(* IEC 61131-3 sources: TBEN-L5-PLC-11/src/st, 44 files *)

(* ---- E_IolAccess.st ---- *)
{attribute 'qualified_only'}
// Quyền truy cập tham số theo IODD (accessRights)
TYPE E_IolAccess :
(
    RO := 0,
    WO := 1,
    RW := 2
) INT;
END_TYPE

(* ---- E_IolCallState.st ---- *)
{attribute 'qualified_only'}
// Trạng thái state machine IOL_CALL của FB_IolMaster
TYPE E_IolCallState :
(
    IDLE      := 0,   // rảnh, chờ request trong FIFO
    WRITE_REQ := 1,   // WRREC khung IOL_CALL vào record CAP 0xB400
    RETRY_WR  := 2,   // master báo bận -> chờ rồi ghi lại
    READ_WAIT := 3,   // REQ đã hạ, chờ trước khi RDREC phản hồi
    READ_REQ  := 4,   // RDREC đọc phản hồi + kiểm khung
    DONE      := 5,   // trả kết quả cho client (1 chu kỳ)
    ERROR     := 6,   // trả lỗi cho client (1 chu kỳ)
    TIMEOUT   := 7,   // quá hạn: hạ REQ, chờ transport hết BUSY
    STUCK     := 8    // transport kẹt BUSY > 1 s, chỉ thoát bằng xReset
) INT;
END_TYPE

(* ---- E_IolCallStep.st ---- *)
{attribute 'qualified_only'}
// Bước handshake của client FB_IolCall
TYPE E_IolCallStep :
(
    IDLE := 0,
    WAIT := 1,    // đã vào hàng đợi master, chờ kết quả
    DONE := 2,
    ERR  := 3
) INT;
END_TYPE

(* ---- E_IolDataType.st ---- *)
{attribute 'qualified_only'}
// Kiểu dữ liệu tham số theo IODD (giá trị trên dây là big-endian)
TYPE E_IolDataType :
(
    U8    := 0,
    U16   := 1,
    U32   := 2,
    I8    := 3,
    I16   := 4,
    I32   := 5,
    STR   := 6,
    OCTET := 7    // record nhiều trường, lớp con tự tách (vd Limit index 64)
) INT;
END_TYPE

(* ---- E_IolDevJob.st ---- *)
{attribute 'qualified_only'}
// Loại việc ISDU đang chạy trong FB_IolDevBase
TYPE E_IolDevJob :
(
    NONE     := 0,
    IDENT    := 1,  // đọc index 16..24
    PARAM_RD := 2,  // đọc 1 tham số trong bảng
    PARAM_WR := 3,  // ghi 1 tham số trong bảng
    CUSTOM   := 4   // ISDU tự do của lớp con (system command, event list...)
) INT;
END_TYPE

(* ---- E_IolDevSeq.st ---- *)
{attribute 'qualified_only'}
// Bước trình tự gọi ISDU trong FB_IolDevBase
TYPE E_IolDevSeq :
(
    IDLE    := 0,   // chọn việc tiếp theo
    RUN     := 1,   // FB_IolCall đang chạy
    RELEASE := 2    // hạ Execute, chờ FB_IolCall về IDLE
) INT;
END_TYPE

(* ---- E_IolErrSource.st ---- *)
{attribute 'qualified_only'}
// Nguồn lỗi của 1 lần gọi IO-Link, để HMI biết lỗi nằm ở tầng nào
TYPE E_IolErrSource :
(
    NONE         := 0,
    PNIO         := 1,    // RDREC/WRREC trả STATUS lỗi (hoặc transport chưa cấu hình)
    IOL_MASTER   := 2,    // AL1100 báo IOL_M_ErrorCode
    IOL_DEVICE   := 3,    // cảm biến báo lỗi ISDU 0x80xx
    TIMEOUT      := 4,
    PARAM        := 5,    // tham số yêu cầu sai, không gửi đi
    LOCK         := 6,    // hết chỗ hàng đợi / không đăng ký được / bị reset
    FRAME        := 7,    // khung phản hồi sai
    NO_DEVICE    := 8,    // PQI.DA = 0: port không có thiết bị
    WRITE_LOCKED := 9,    // ghi bị khoá (chưa bật xMaintEnable)
    RANGE        := 10    // giá trị đặt ngoài dải IODD, chặn trước khi gửi
) INT;
END_TYPE

(* ---- E_IolEvtType.st ---- *)
{attribute 'qualified_only'}
// Loại event IO-Link (= bit 5..4 của EventQualifier)
TYPE E_IolEvtType :
(
    NOTIFICATION := 1,
    WARNING      := 2,
    ERROR        := 3
) INT;
END_TYPE

(* ---- E_IolService.st ---- *)
{attribute 'qualified_only'}
// Giá trị byte Control của khung IOL_CALL (request)
TYPE E_IolService :
(
    WRITE := 2,   // ISDU write
    READ  := 3    // ISDU read
) USINT;
END_TYPE

(* ---- E_O5D150_Param.st ---- *)
{attribute 'qualified_only'}
// Vị trí tham số trong bảng GVL_O5D150_Def.aParamDef (không phải IO-Link index)
TYPE E_O5D150_Param :
(
    SP1       := 0,   // index 60 sub 1
    CFG_LOGIC := 1,   // index 61 sub 1
    LIMITS    := 2,   // index 64 (min, max) - không đặt tên LIMIT vì trùng hàm chuẩn
    ALIGN     := 3,   // index 69
    LASER     := 4,   // index 80
    DISPLAY   := 5,   // index 96
    KEYLOCK   := 6,   // index 100
    DFO       := 7,   // index 74
    DS        := 8,   // index 76
    DR        := 9    // index 78
) INT;
END_TYPE

(* ---- ST_HMI_O5D150.st ---- *)
// Giao tiếp HMI <-> FB_Dev_O5D150 (lệnh: HMI đặt TRUE, PRG_IOLink tự xoá)
TYPE ST_HMI_O5D150 :
STRUCT
    // --- Lệnh ---
    xCmdReadAll      : BOOL;
    xCmdReadIdent    : BOOL;
    xCmdWriteSP1     : BOOL;          // ghi uiSetSP1 (cần xMaintEnable)
    xCmdWriteLogic   : BOOL;
    xCmdWriteLaser   : BOOL;
    xCmdWriteDisplay : BOOL;
    xCmdTestEvt1On   : BOOL;          // System Command 240 (cần xMaintEnable)
    xCmdTestEvt1Off  : BOOL;          // 241
    xCmdTestEvt2On   : BOOL;          // 242
    xCmdTestEvt2Off  : BOOL;          // 243
    xCmdReadEvents   : BOOL;          // đọc index 37 ngay (thử lại cả khi đã báo không hỗ trợ)
    xCmdResetErr     : BOOL;
    xAlignMode       : BOOL;          // giữ TRUE: đọc Align (69) chu kỳ chậm

    // --- Giá trị đặt ---
    uiSetSP1         : UINT := 100;   // cm, 5..200
    usiSetLogic      : USINT;         // 0 NO, 1 NC
    usiSetLaser      : USINT := 1;    // 0 Off, 1 On
    usiSetDisplay    : USINT := 1;    // 0 Off, 1 On, 2 Rotated

    // --- Process data ---
    uiDistance_cm    : UINT;
    rDistance_m      : REAL;
    xOut1            : BOOL;
    xPdValid         : BOOL;
    xOutOfRange      : BOOL;
    xPQ              : BOOL;
    xDA              : BOOL;
    xDE              : BOOL;

    // --- Tham số đọc về ---
    uiSP1            : UINT;
    usiLogic         : USINT;
    uiLimitMin_cm    : UINT;
    uiLimitMax_cm    : UINT;
    usiAlign         : USINT;         // %
    usiLaser         : USINT;
    usiDisplay       : USINT;
    xParamValid      : BOOL;          // SP1 đọc được lần gần nhất

    // --- Nhận dạng ---
    sVendor          : STRING(64);
    sProduct         : STRING(64);
    sSerial          : STRING(64);
    sFwRev           : STRING(64);

    // --- Event ---
    axEvtActive      : ARRAY[0..GVL_O5D150_Def.iEVT_COUNT - 1] OF BOOL;   // theo GVL_O5D150_Def.aEvtDef
    uiEvtCount       : UINT;
    wUnknownEvt      : WORD;
    xEvtListNotSupported : BOOL;

    // --- Trạng thái / lỗi ---
    xBusy            : BOOL;
    xError           : BOOL;          // lỗi gần nhất (giữ tới xCmdResetErr)
    uiDevErr         : UINT;
    wsErrText        : WSTRING(80);
    xWriteLocked     : BOOL;          // = NOT xMaintEnable
END_STRUCT
END_TYPE

(* ---- ST_IolEventDef.st ---- *)
// Định nghĩa 1 event của device (từ IODD)
TYPE ST_IolEventDef :
STRUCT
    wCode  : WORD;
    sName  : STRING(12);        // tên ngắn trên màn hình cảm biến
    wsText : WSTRING(48);       // mô tả cho HMI
    eType  : E_IolEvtType;
END_STRUCT
END_TYPE

(* ---- ST_IolIdent.st ---- *)
// Thông tin nhận dạng chuẩn IO-Link (index 16..24)
TYPE ST_IolIdent :
STRUCT
    sVendorName  : STRING(64);   // 16
    sVendorText  : STRING(64);   // 17
    sProductName : STRING(64);   // 18
    sProductId   : STRING(64);   // 19
    sProductText : STRING(64);   // 20
    sSerialNo    : STRING(64);   // 21
    sHwRev       : STRING(64);   // 22
    sFwRev       : STRING(64);   // 23
    sAppTag      : STRING(64);   // 24
END_STRUCT
END_TYPE

(* ---- ST_IolParamDef.st ---- *)
// Định nghĩa 1 tham số lấy từ IODD (bảng hằng trong GVL_<Model>_Def)
TYPE ST_IolParamDef :
STRUCT
    sName       : STRING(24);                  // tên theo IODD
    uiIndex     : UINT;
    usiSubindex : USINT;                       // 0 = cả index
    eType       : E_IolDataType;
    eAccess     : E_IolAccess;
    diMin       : DINT;                        // dải hợp lệ khi ghi (raw = đơn vị kỹ thuật)
    diMax       : DINT;
    diDefault   : DINT;
    sUnit       : STRING(8);
    xInReadAll  : BOOL := TRUE;                // có đọc trong ReadAll không
END_STRUCT
END_TYPE

(* ---- ST_IolParamVal.st ---- *)
// Giá trị runtime của 1 tham số (không RETAIN: nguồn thật là cảm biến)
TYPE ST_IolParamVal :
STRUCT
    diRaw  : DINT;      // giá trị đọc về gần nhất
    xValid : BOOL;      // lần đọc gần nhất thành công
    uiErr  : UINT;      // 0x80xx = lỗi device, 0xFFnn = lỗi nội bộ (nn = E_IolErrSource)
    diSet  : DINT;      // giá trị đang chờ ghi
    xDirty : BOOL;      // TRUE từ lúc yêu cầu ghi tới khi ghi xong
END_STRUCT
END_TYPE

(* ---- ST_IolPortDiag.st ---- *)
// Port Qualifier (PQI) AL1100 đã giải mã - bit theo GSDML ifm AL1100
TYPE ST_IolPortDiag :
STRUCT
    bPQI : BYTE;
    xDI4 : BOOL;   // bit0 trạng thái chân 4 (DI)
    xDI2 : BOOL;   // bit1 trạng thái chân 2 (DI)
    xNP  : BOOL;   // bit2
    xSV  : BOOL;   // bit3
    xDA  : BOOL;   // bit4 Device Available
    xDC  : BOOL;   // bit5
    xDE  : BOOL;   // bit6 Device Error
    xPQ  : BOOL;   // bit7 Port Qualifier: PDin hợp lệ
END_STRUCT
END_TYPE

(* ---- ST_IolRequest.st ---- *)
// 1 request ISDU gửi qua master
TYPE ST_IolRequest :
STRUCT
    usiPort     : USINT;                                   // 0 = master, 1..4 = port
    eService    : E_IolService := E_IolService.READ;
    uiIndex     : UINT;
    usiSubindex : USINT;                                   // 0 = cả index
    uiLen       : UINT;                                    // số byte dữ liệu ghi (READ = 0)
    abData      : ARRAY[0..GVL_IolConst.uiMAX_DATA - 1] OF BYTE;
END_STRUCT
END_TYPE

(* ---- ST_IolResult.st ---- *)
// Kết quả 1 request ISDU master trả cho client
TYPE ST_IolResult :
STRUCT
    xError         : BOOL;
    eErrSource     : E_IolErrSource;
    dwPnioStatus   : DWORD;                                // STATUS RDREC/WRREC
    uiIolMasterErr : UINT;                                 // IOL_M_ErrorCode
    uiIolDevErr    : UINT;                                 // lỗi ISDU device 0x80xx
    uiLen          : UINT;                                 // số byte dữ liệu đọc về
    abData         : ARRAY[0..GVL_IolConst.uiMAX_DATA - 1] OF BYTE;
END_STRUCT
END_TYPE

(* ---- ST_MockParam.st ---- *)
// 1 index trong bảng dữ liệu giả lập của FB_MockRecordAccess
TYPE ST_MockParam :
STRUCT
    uiIndex : UINT;
    eAccess : E_IolAccess;
    uiLen   : UINT;                      // số byte của cả index
    abData  : ARRAY[0..63] OF BYTE;      // big-endian như trên dây
END_STRUCT
END_TYPE

(* ---- ST_O5D150_PdIn.st ---- *)
// PDin O5D150 đã giải mã
TYPE ST_O5D150_PdIn :
STRUCT
    wRaw          : WORD;     // word PDin ghép big-endian
    uiDistance_cm : UINT;     // giữ giá trị cũ khi PD không hợp lệ
    rDistance_m   : REAL;
    xOut1         : BOOL;     // FALSE (fail-safe) khi PD không hợp lệ
    xPdValid      : BOOL;     // PQ AND DA
    xOutOfRange   : BOOL;     // ngoài 5..200 cm (không có vật / quá gần)
END_STRUCT
END_TYPE

(* ---- ST_O5D150_PdLayout.st ---- *)
// Bố cục PDin O5D150 (16 bit, big-endian) - tách thành hằng để sửa theo IODD mà không đổi logic
TYPE ST_O5D150_PdLayout :
STRUCT
    usiOut1Bit       : USINT;      // bit OUT1 trong word PDin
    usiDistBitOffset : USINT;      // bit bắt đầu của Distance
    wDistMask        : WORD;       // mặt nạ sau khi dịch (12 bit = 16#0FFF)
    uiDistMin        : UINT;       // dải đo hợp lệ [cm]
    uiDistMax        : UINT;
    rGradient        : REAL;       // m / digit
END_STRUCT
END_TYPE

(* ---- GVL_HMI_IOL.st ---- *)
{attribute 'qualified_only'}
// Giao tiếp HMI cho IO-Link (tách khỏi GVL_HMI của trình tự đèn DXP)
VAR_GLOBAL
    xMaintEnable    : BOOL;                 // cho phép ghi tham số / System Command (khoá mặc định)
    xCmdResetMaster : BOOL;                 // xoá hàng đợi / thoát STUCK (chỉ khi xMaintEnable)
    stO5D150        : ST_HMI_O5D150;        // O5D150 port 1

    // --- Trạng thái master AL1100 ---
    eMasterState    : E_IolCallState;
    udiCallCount    : UDINT;
    udiErrCount     : UDINT;
    xSimMode        : BOOL;                 // bản sao GVL_IolSys.xSimMode để hiển thị

    // --- Alarm (bit) ---
    xAlmP1_NoDevice   : BOOL;               // PQI.DA = 0 > 2 s
    xAlmP1_PdInvalid  : BOOL;               // DA = 1 nhưng PQ = 0 > 1 s
    xAlmP1_DevErr     : BOOL;               // PQI.DE
    xAlmP1_EvtError   : BOOL;               // có event loại ERROR đang active
    xAlmIolCallErr    : BOOL;               // lần gọi ISDU gần nhất lỗi
    xAlmMasterStuck   : BOOL;               // master kẹt, cần xCmdResetMaster
    xAlarmAny         : BOOL;               // OR các alarm mức Lỗi
    xWarningAny       : BOOL;               // OR các cảnh báo
END_VAR

(* ---- GVL_IO.st ---- *)
// Ngõ vào/ra DXP của TBEN-L5-PLC-11 (map trong Local_IO > DXP > I/O Mapping)
// Đầu nối: C4 = Ch8/Ch9, C5 = Ch10/Ch11, C6 = Ch12/Ch13, C7 = Ch14/Ch15
VAR_GLOBAL
    xQ_Ch8  : BOOL;   // ngõ ra DXP Ch8  (C4)
    xQ_Ch9  : BOOL;   // ngõ ra DXP Ch9  (C4)
    xQ_Ch10 : BOOL;   // ngõ ra DXP Ch10 (C5)
    xQ_Ch11 : BOOL;   // ngõ ra DXP Ch11 (C5)
    xQ_Ch12 : BOOL;   // ngõ ra DXP Ch12 (C6)
    xQ_Ch13 : BOOL;   // ngõ ra DXP Ch13 (C6)
    xQ_Ch14 : BOOL;   // ngõ ra DXP Ch14 (C7)
    xQ_Ch15 : BOOL;   // ngõ ra DXP Ch15 (C7)

    xI_Ch8  : BOOL;   // đọc lại mức tín hiệu DXP Ch8
    xI_Ch9  : BOOL;   // đọc lại mức tín hiệu DXP Ch9
    xI_Ch10 : BOOL;   // đọc lại mức tín hiệu DXP Ch10
    xI_Ch11 : BOOL;   // đọc lại mức tín hiệu DXP Ch11
    xI_Ch12 : BOOL;   // đọc lại mức tín hiệu DXP Ch12
    xI_Ch13 : BOOL;   // đọc lại mức tín hiệu DXP Ch13
    xI_Ch14 : BOOL;   // đọc lại mức tín hiệu DXP Ch14
    xI_Ch15 : BOOL;   // đọc lại mức tín hiệu DXP Ch15

    // IO-Link master ifm AL1100 (PROFINET), port 1 = O5D150.
    // TODO PROFINET: map 2 biến này vào Input data / PQI của submodule Port 1 khi thêm AL1100; hiện là biến thường để Write/Force trên Simulation.
    abAL1_P1_In : ARRAY[0..1] OF BYTE;   // PDin O5D150 big-endian: byte 0 = MSB (Distance bit 15..4, OUT1 bit 0)
    bAL1_P1_PQI : BYTE;                  // Port Qualifier: bit7 PQ, bit6 DE, bit5 DC, bit4 DA (16#90 = PQ + DA)
END_VAR

(* ---- GVL_IolConst.st ---- *)
{attribute 'qualified_only'}
// Hằng số IO-Link Call qua PROFINET (spec PNO "IO-Link Integration for PROFINET")
VAR_GLOBAL CONSTANT
    // --- Khung IOL_CALL (record CAP) ---
    uiCAP_INDEX        : UINT  := 16#B400;   // record index CAP; CommFB.INDEX là INT -> truyền UINT_TO_INT (bit pattern giữ nguyên)
    usiEXT_FUNC_NUM    : USINT := 16#08;     // byte 0 khung IOL_CALL
    uiFI_INDEX         : UINT  := 16#FE4A;   // function index IOL_CALL (65098)
    usiCTRL_RELEASE    : USINT := 0;
    usiCTRL_WRITE      : USINT := 2;
    usiCTRL_READ       : USINT := 3;
    usiCTRL_ERROR      : USINT := 16#80;     // Control phản hồi lỗi - cần đối chiếu manual AL1100
    uiHDR_LEN          : UINT  := 8;         // header khung IOL_CALL
    uiMAX_DATA         : UINT  := 232;       // dữ liệu ISDU tối đa trong 1 IOL_CALL
    uiMAX_REC          : UINT  := 240;       // MLEN của RDREC = header + data

    // --- Vị trí AL1100 / thiết bị ---
    usiAL1_SLOT        : USINT := 1;         // submodule "IO-Link Master" (giả định, dự phòng slot 0/subslot 1)
    usiAL1_SUBSLOT_CAP : USINT := 1;
    usiPORT_O5D150     : USINT := 1;         // O5D150 cắm port X01 - đổi port tại đây

    // --- Thời gian / giới hạn ---
    tCALL_TIMEOUT      : TIME  := T#5S;      // tổng thời gian 1 request trong master
    tRETRY_DELAY       : TIME  := T#20MS;    // chờ giữa các lần RDREC khi master còn bận
    iMAX_RETRY         : INT   := 100;
    iQUEUE_SIZE        : INT   := 16;        // số client tối đa trên 1 master
    iMAX_PARAM         : INT   := 32;        // số tham số tối đa trong bảng của 1 device

    // --- Mã lỗi ISDU hay dùng ---
    uiERR_IDX_NA       : UINT  := 16#8011;   // index không tồn tại
    uiERR_SUBIDX_NA    : UINT  := 16#8012;
    uiERR_ACCESS       : UINT  := 16#8023;
    uiERR_RANGE        : UINT  := 16#8030;

    // --- STATUS nội bộ (không phải mã PNIO thật) ---
    dwSTAT_NOT_CONFIGURED : DWORD := 16#FFFF0001;  // FB_PnRecordAccess còn là khung, chưa có PN Controller
    dwSTAT_NO_TRANSPORT   : DWORD := 16#FFFF0002;  // master chưa được gán itfRec
END_VAR

(* ---- GVL_IolSys.st ---- *)
{attribute 'qualified_only'}
// Instance master + transport IO-Link (gọi trong PRG_IOLink / MainTask)
VAR_GLOBAL
    xSimMode  : BOOL := TRUE;              // TRUE = dùng mock (Simulation). Đặt FALSE sau khi có PROFINET thật.
    fbMockAL1 : FB_MockRecordAccess;       // giả lập AL1100 + O5D150
    fbPnAL1   : FB_PnRecordAccess;         // transport PROFINET thật (hiện là khung)
    fbAL1     : FB_IolMaster;              // master AL1100: khoá + hàng đợi IOL_CALL
END_VAR

(* ---- GVL_O5D150_Def.st ---- *)
{attribute 'qualified_only'}
// Bảng hằng O5D150 lấy từ IODD ifm-000174-20210526-IODD1.1.xml (vendor 310, device 372)
VAR_GLOBAL CONSTANT
    uiPDIN_LEN   : UINT := 2;
    stPdLayout   : ST_O5D150_PdLayout := (usiOut1Bit := 0, usiDistBitOffset := 4, wDistMask := 16#0FFF,
                                          uiDistMin := 5, uiDistMax := 200, rGradient := 0.01);

    iPARAM_COUNT : INT := 10;   // = số phần tử E_O5D150_Param
    aParamDef    : ARRAY[0..9] OF ST_IolParamDef := [
        (sName := 'SP1',     uiIndex := 60,  usiSubindex := 1, eType := E_IolDataType.U16, eAccess := E_IolAccess.RW, diMin := 5, diMax := 200,  diDefault := 100, sUnit := 'cm', xInReadAll := TRUE),
        (sName := 'Logic',   uiIndex := 61,  usiSubindex := 1, eType := E_IolDataType.U8,  eAccess := E_IolAccess.RW, diMin := 0, diMax := 1,    diDefault := 0,   sUnit := '',   xInReadAll := TRUE),
        (sName := 'Limit',   uiIndex := 64,  usiSubindex := 0, eType := E_IolDataType.U32, eAccess := E_IolAccess.RO, diMin := 0, diMax := 0,    diDefault := 0,   sUnit := 'cm', xInReadAll := TRUE),
        (sName := 'Align',   uiIndex := 69,  usiSubindex := 0, eType := E_IolDataType.U8,  eAccess := E_IolAccess.RO, diMin := 0, diMax := 100,  diDefault := 0,   sUnit := '%',  xInReadAll := TRUE),
        (sName := 'Laser',   uiIndex := 80,  usiSubindex := 0, eType := E_IolDataType.U8,  eAccess := E_IolAccess.RW, diMin := 0, diMax := 1,    diDefault := 1,   sUnit := '',   xInReadAll := TRUE),
        (sName := 'Display', uiIndex := 96,  usiSubindex := 0, eType := E_IolDataType.U8,  eAccess := E_IolAccess.RW, diMin := 0, diMax := 2,    diDefault := 1,   sUnit := '',   xInReadAll := TRUE),
        (sName := 'KeyLock', uiIndex := 100, usiSubindex := 0, eType := E_IolDataType.U8,  eAccess := E_IolAccess.RW, diMin := 0, diMax := 1,    diDefault := 1,   sUnit := '',   xInReadAll := TRUE),
        (sName := 'dFO',     uiIndex := 74,  usiSubindex := 0, eType := E_IolDataType.U16, eAccess := E_IolAccess.RW, diMin := 0, diMax := 2000, diDefault := 0,   sUnit := '',   xInReadAll := TRUE),
        (sName := 'dS',      uiIndex := 76,  usiSubindex := 0, eType := E_IolDataType.U16, eAccess := E_IolAccess.RW, diMin := 0, diMax := 2000, diDefault := 0,   sUnit := '',   xInReadAll := TRUE),
        (sName := 'dr',      uiIndex := 78,  usiSubindex := 0, eType := E_IolDataType.U16, eAccess := E_IolAccess.RW, diMin := 0, diMax := 2000, diDefault := 0,   sUnit := '',   xInReadAll := TRUE)
    ];

    // --- System Command (index 2, UINT8, write only) ---
    uiIDX_SYS_CMD        : UINT  := 2;
    usiSC_FACTORY_RESET  : USINT := 130;
    usiSC_TEST_EVT1_ON   : USINT := 240;   // Test Event 0x8DFE appear
    usiSC_TEST_EVT1_OFF  : USINT := 241;   // Test Event 0x8DFE disappear
    usiSC_TEST_EVT2_ON   : USINT := 242;   // Test Event 0x8DFF appear
    usiSC_TEST_EVT2_OFF  : USINT := 243;   // Test Event 0x8DFF disappear

    // --- Event (Detailed Device Status index 37: 3 byte/entry; IODD không khai báo -> có thể trả 0x8011) ---
    uiIDX_EVT_LIST : UINT := 37;
    iEVT_COUNT     : INT  := 8;
    aEvtDef        : ARRAY[0..7] OF ST_IolEventDef := [
        (wCode := 16#4220, sName := 'TEMP', wsText := "Quá nhiệt thiết bị",                 eType := E_IolEvtType.WARNING),
        (wCode := 16#8CB0, sName := 'nEA',  wsText := "Cảnh báo: vật quá gần",              eType := E_IolEvtType.WARNING),
        (wCode := 16#8CB1, sName := 'fAr',  wsText := "Cảnh báo: vật quá xa",               eType := E_IolEvtType.WARNING),
        (wCode := 16#8CB4, sName := '+',    wsText := "Lỗi: cường độ phản xạ quá lớn",     eType := E_IolEvtType.ERROR),
        (wCode := 16#8CB5, sName := '-',    wsText := "Lỗi: không có vật / tín hiệu",       eType := E_IolEvtType.ERROR),
        (wCode := 16#8CA4, sName := 'ErP',  wsText := "Cảnh báo: sai lệch tính hợp lý",     eType := E_IolEvtType.WARNING),
        (wCode := 16#8DFE, sName := 'TEST1', wsText := "Sự kiện thử 1 (System Command 240)", eType := E_IolEvtType.NOTIFICATION),
        (wCode := 16#8DFF, sName := 'TEST2', wsText := "Sự kiện thử 2 (System Command 242)", eType := E_IolEvtType.NOTIFICATION)
    ];
END_VAR

(* ---- ITF_IolRecordAccess.st ---- *)
// Ghi record (WRREC). Trả TRUE khi đã kết thúc (xDone hoặc xError).
METHOD Write : BOOL
VAR_INPUT
    xReq   : BOOL;
    dwId   : DWORD;                 // ID submodule (CommFB.SUBSLOT_ID), mock bỏ qua
    iIndex : INT;                   // record index (0xB400 truyền dạng INT)
    iLen   : INT;                   // số byte ghi
    pData  : POINTER TO BYTE;
END_VAR
VAR_OUTPUT
    xDone    : BOOL;
    xBusy    : BOOL;
    xError   : BOOL;
    dwStatus : DWORD;               // STATUS PNIO 4 byte
END_VAR

// Đọc record (RDREC). Trả TRUE khi đã kết thúc (xValid hoặc xError).
METHOD Read : BOOL
VAR_INPUT
    xReq   : BOOL;
    dwId   : DWORD;
    iIndex : INT;
    iMLen  : INT;                   // kích thước buffer nhận
    pData  : POINTER TO BYTE;
END_VAR
VAR_OUTPUT
    xValid   : BOOL;
    xBusy    : BOOL;
    xError   : BOOL;
    dwStatus : DWORD;
    iLen     : INT;                 // số byte nhận được
END_VAR

// Trừu tượng hoá đọc/ghi record PROFINET (CommFB.WRREC/RDREC thật hoặc mock Simulation)
// Quy ước như CommFB: giữ xReq = TRUE tới khi có kết quả, hạ xReq ít nhất 1 lần gọi trước request mới; gọi mỗi chu kỳ đúng 1 lần.
INTERFACE ITF_IolRecordAccess

(* ---- F_IolBytesToStr.st ---- *)
// Chuyển StringT IO-Link (không có ký tự kết thúc) thành STRING, cắt ở 64 ký tự
FUNCTION F_IolBytesToStr : STRING(64)
VAR_INPUT
    pBuf  : POINTER TO BYTE;
    uiLen : UINT;
END_VAR
VAR
    sTmp : STRING(64);
    pDst : POINTER TO BYTE;
    i    : UINT;
    n    : UINT;
END_VAR

(*---IMPL---*)
sTmp := '';
IF pBuf <> 0 THEN
    n := MIN(uiLen, 64);
    pDst := ADR(sTmp);
    i := 0;
    WHILE i < n DO
        IF pBuf[i] = 0 THEN          // device có thể đệm 0 ở cuối
            EXIT;
        END_IF
        pDst[i] := pBuf[i];
        i := i + 1;
    END_WHILE
    pDst[i] := 0;
END_IF
F_IolBytesToStr := sTmp;

(* ---- F_IolErrText.st ---- *)
// Mã lỗi IO-Link Call -> chuỗi hiển thị HMI
FUNCTION F_IolErrText : WSTRING(80)
VAR_INPUT
    eSrc       : E_IolErrSource;
    uiMasterEr : UINT;        // IOL_M_ErrorCode
    uiDevErr   : UINT;        // lỗi ISDU 0x80xx
    dwPnio     : DWORD;       // STATUS RDREC/WRREC
END_VAR

(*---IMPL---*)
CASE eSrc OF
    E_IolErrSource.NONE:
        F_IolErrText := "OK";

    E_IolErrSource.PNIO:
        IF dwPnio = GVL_IolConst.dwSTAT_NOT_CONFIGURED THEN
            F_IolErrText := "PROFINET chưa cấu hình (FB_PnRecordAccess còn là khung)";
        ELSIF dwPnio = GVL_IolConst.dwSTAT_NO_TRANSPORT THEN
            F_IolErrText := "Master chưa gán transport (itfRec)";
        ELSIF F_IolIsPnioBusy(dwPnio) THEN
            F_IolErrText := "AL1100 bận quá số lần thử lại";
        ELSE
            F_IolErrText := "Lỗi đọc/ghi record PROFINET (xem dwPnioStatus)";
        END_IF

    E_IolErrSource.IOL_MASTER:
        CASE uiMasterEr OF
            16#7000: F_IolErrText := "Master: xung đột IOL_CALL";
            16#7001: F_IolErrText := "Master: khung IOL_CALL sai";
            16#7002: F_IolErrText := "Master: port đang bị khoá";
            16#8000: F_IolErrText := "Master: timeout";
            16#8001: F_IolErrText := "Master: số port không hợp lệ";
            16#8002: F_IolErrText := "Master: chế độ port không phải IO-Link";
            16#8003: F_IolErrText := "Master: độ dài không hợp lệ";
            16#8004: F_IolErrText := "Master: lỗi truyền thông với thiết bị";
        ELSE
            F_IolErrText := "Master: lỗi khác (xem uiIolMasterErr)";
        END_CASE

    E_IolErrSource.IOL_DEVICE:
        CASE uiDevErr OF
            16#8000: F_IolErrText := "Thiết bị: lỗi ứng dụng";
            16#8011: F_IolErrText := "Thiết bị: index không tồn tại";
            16#8012: F_IolErrText := "Thiết bị: subindex không tồn tại";
            16#8020, 16#8021, 16#8022:
                     F_IolErrText := "Thiết bị: dịch vụ tạm thời không sẵn sàng";
            16#8023: F_IolErrText := "Thiết bị: từ chối truy cập";
            16#8030: F_IolErrText := "Thiết bị: giá trị ngoài dải";
            16#8031: F_IolErrText := "Thiết bị: giá trị vượt giới hạn trên";
            16#8032: F_IolErrText := "Thiết bị: giá trị dưới giới hạn dưới";
            16#8033: F_IolErrText := "Thiết bị: dữ liệu quá dài";
            16#8034: F_IolErrText := "Thiết bị: dữ liệu quá ngắn";
            16#8035: F_IolErrText := "Thiết bị: chức năng không hỗ trợ";
            16#8036: F_IolErrText := "Thiết bị: chức năng tạm không sẵn sàng";
            16#8040: F_IolErrText := "Thiết bị: bộ tham số không hợp lệ";
            16#8041: F_IolErrText := "Thiết bị: bộ tham số không nhất quán";
            16#8082: F_IolErrText := "Thiết bị: ứng dụng chưa sẵn sàng";
        ELSE
            F_IolErrText := "Thiết bị: lỗi khác (xem uiIolDevErr)";
        END_CASE

    E_IolErrSource.TIMEOUT:
        F_IolErrText := "Quá thời gian chờ phản hồi";
    E_IolErrSource.PARAM:
        F_IolErrText := "Tham số yêu cầu sai, không gửi";
    E_IolErrSource.LOCK:
        F_IolErrText := "Hàng đợi master đầy hoặc đã bị reset";
    E_IolErrSource.FRAME:
        F_IolErrText := "Khung phản hồi IOL_CALL sai";
    E_IolErrSource.NO_DEVICE:
        F_IolErrText := "Port không có thiết bị (PQI.DA = 0)";
    E_IolErrSource.WRITE_LOCKED:
        F_IolErrText := "Ghi bị khoá: chưa bật xMaintEnable";
    E_IolErrSource.RANGE:
        F_IolErrText := "Giá trị đặt ngoài dải IODD, không gửi";
ELSE
    F_IolErrText := "Lỗi không xác định";
END_CASE

(* ---- F_IolGetR32BE.st ---- *)
// Đọc Float32T IO-Link (IEEE754 big-endian): chép bit pattern, không đổi số học
FUNCTION F_IolGetR32BE : REAL
VAR_INPUT
    pBuf  : POINTER TO BYTE;
    uiOff : UINT;
END_VAR
VAR
    dwTmp : DWORD;
    pR    : POINTER TO REAL;
END_VAR

(*---IMPL---*)
dwTmp := F_IolGetU32BE(pBuf, uiOff);
pR := ADR(dwTmp);
F_IolGetR32BE := pR^;

(* ---- F_IolGetU16BE.st ---- *)
// Đọc UINT big-endian (IO-Link/PROFINET) từ buffer byte - TBEN là ARM little-endian nên không ép kiểu trực tiếp
FUNCTION F_IolGetU16BE : UINT
VAR_INPUT
    pBuf  : POINTER TO BYTE;
    uiOff : UINT;               // vị trí byte MSB
END_VAR

(*---IMPL---*)
IF pBuf = 0 THEN
    F_IolGetU16BE := 0;
    RETURN;
END_IF
F_IolGetU16BE := WORD_TO_UINT(SHL(BYTE_TO_WORD(pBuf[uiOff]), 8) OR BYTE_TO_WORD(pBuf[uiOff + 1]));

(* ---- F_IolGetU32BE.st ---- *)
// Đọc 4 byte big-endian thành DWORD
FUNCTION F_IolGetU32BE : DWORD
VAR_INPUT
    pBuf  : POINTER TO BYTE;
    uiOff : UINT;
END_VAR

(*---IMPL---*)
IF pBuf = 0 THEN
    F_IolGetU32BE := 0;
    RETURN;
END_IF
F_IolGetU32BE := SHL(UINT_TO_DWORD(F_IolGetU16BE(pBuf, uiOff)), 16) OR UINT_TO_DWORD(F_IolGetU16BE(pBuf, uiOff + 2));

(* ---- F_IolIsPnioBusy.st ---- *)
// TRUE nếu STATUS RDREC/WRREC là "state conflict" (B5) hoặc "resource busy" (C3) -> master chưa xong, được retry
FUNCTION F_IolIsPnioBusy : BOOL
VAR_INPUT
    dwStatus : DWORD;          // ErrorCode, ErrorDecode, ErrorCode1, ErrorCode2 (byte cao -> thấp)
END_VAR
VAR
    bCode1 : BYTE;
END_VAR

(*---IMPL---*)
bCode1 := DWORD_TO_BYTE(SHR(dwStatus, 8));
F_IolIsPnioBusy := (bCode1 = 16#B5) OR (bCode1 = 16#C3);

(* ---- F_IolSetR32BE.st ---- *)
// Ghi REAL dạng Float32T big-endian
FUNCTION F_IolSetR32BE : BOOL
VAR_INPUT
    pBuf  : POINTER TO BYTE;
    uiOff : UINT;
    rVal  : REAL;
END_VAR
VAR
    pDw : POINTER TO DWORD;
END_VAR

(*---IMPL---*)
pDw := ADR(rVal);
F_IolSetR32BE := F_IolSetU32BE(pBuf, uiOff, pDw^);

(* ---- F_IolSetU16BE.st ---- *)
// Ghi UINT big-endian vào buffer byte; FALSE nếu pBuf = 0
FUNCTION F_IolSetU16BE : BOOL
VAR_INPUT
    pBuf  : POINTER TO BYTE;
    uiOff : UINT;
    uiVal : UINT;
END_VAR

(*---IMPL---*)
IF pBuf = 0 THEN
    F_IolSetU16BE := FALSE;
    RETURN;
END_IF
pBuf[uiOff]     := WORD_TO_BYTE(SHR(UINT_TO_WORD(uiVal), 8));
pBuf[uiOff + 1] := UINT_TO_BYTE(uiVal);
F_IolSetU16BE := TRUE;

(* ---- F_IolSetU32BE.st ---- *)
// Ghi DWORD big-endian (4 byte) vào buffer
FUNCTION F_IolSetU32BE : BOOL
VAR_INPUT
    pBuf  : POINTER TO BYTE;
    uiOff : UINT;
    dwVal : DWORD;
END_VAR

(*---IMPL---*)
IF pBuf = 0 THEN
    F_IolSetU32BE := FALSE;
    RETURN;
END_IF
F_IolSetU16BE(pBuf, uiOff, DWORD_TO_UINT(SHR(dwVal, 16)));
F_IolSetU16BE(pBuf, uiOff + 2, DWORD_TO_UINT(dwVal));
F_IolSetU32BE := TRUE;

(* ---- FB_Dev_O5D150.st ---- *)
// Cảm biến khoảng cách laser ifm O5D150 (IODD vendor 310 / device 372, IO-Link 1.1, PDin 16 bit, không PDout).
// 1) Cyclic: giải mã PDin + PQI.  2) Event: Test Event qua System Command, đọc danh sách event index 37.
// 3) Acyclic: SP1, Logic, Limit, Align, Laser, Display... theo bảng GVL_O5D150_Def.aParamDef.
FUNCTION_BLOCK FB_Dev_O5D150 EXTENDS FB_IolDevBase
VAR_INPUT
    abPdIn           : ARRAY[0..1] OF BYTE;    // PDin từ GVL_IO, big-endian
    xAlignMode       : BOOL;                   // TRUE: đọc Align (69) mỗi tAlignPoll
    // --- Lệnh (sườn lên) ---
    xCmdReadAll      : BOOL;
    xCmdReadIdent    : BOOL;
    xCmdWriteSP1     : BOOL;
    xCmdWriteLogic   : BOOL;
    xCmdWriteLaser   : BOOL;
    xCmdWriteDisplay : BOOL;
    xCmdTestEvt1On   : BOOL;
    xCmdTestEvt1Off  : BOOL;
    xCmdTestEvt2On   : BOOL;
    xCmdTestEvt2Off  : BOOL;
    xCmdReadEvents   : BOOL;
    // --- Giá trị đặt ---
    uiSetSP1         : UINT;                   // cm 5..200
    usiSetLogic      : USINT;                  // 0 NO / 1 NC
    usiSetLaser      : USINT;                  // 0 Off / 1 On
    usiSetDisplay    : USINT;                  // 0 Off / 1 On / 2 Rotated
    tAlignPoll       : TIME := T#500MS;
    tEvtPoll         : TIME := T#5S;           // chu kỳ đọc index 37 khi PD hợp lệ
END_VAR
VAR_OUTPUT
    stPd                 : ST_O5D150_PdIn;
    aVal                 : ARRAY[0..GVL_O5D150_Def.iPARAM_COUNT - 1] OF ST_IolParamVal;   // theo E_O5D150_Param
    uiLimitMin_cm        : UINT;
    uiLimitMax_cm        : UINT;
    axEvtActive          : ARRAY[0..GVL_O5D150_Def.iEVT_COUNT - 1] OF BOOL;   // theo GVL_O5D150_Def.aEvtDef
    xEvtErrorActive      : BOOL;               // có event loại ERROR đang active
    uiEvtCount           : UINT;               // số event đang active (kể cả mã lạ)
    wUnknownEvt          : WORD;               // mã event không có trong bảng (gần nhất)
    xEvtListValid        : BOOL;               // danh sách event đọc được lần gần nhất
    xEvtListNotSupported : BOOL;               // device trả 0x8011 cho index 37 -> ngừng đọc chu kỳ
END_VAR
VAR
    rtReadAll    : R_TRIG;
    rtReadIdent  : R_TRIG;
    rtWrSP1      : R_TRIG;
    rtWrLogic    : R_TRIG;
    rtWrLaser    : R_TRIG;
    rtWrDisplay  : R_TRIG;
    rtEvt1On     : R_TRIG;
    rtEvt1Off    : R_TRIG;
    rtEvt2On     : R_TRIG;
    rtEvt2Off    : R_TRIG;
    rtReadEvt    : R_TRIG;
    tonAlign     : TON;
    tonEvt       : TON;
    usiPendSysCmd: USINT;                      // System Command chờ gửi, 0 = không
    xPendEvtRead : BOOL;
    abCmd        : ARRAY[0..0] OF BYTE;
END_VAR

(*---IMPL---*)
// Nền: PQI, trình tự ISDU, Ident (FB_IolDevBase)
SUPER^();

// ---------- 1. Process data cyclic ----------
DecodePdIn();

// ---------- 2. Lệnh tham số (ghi bị chặn trong RequestWrite nếu chưa bật Maintenance / ngoài dải) ----------
rtReadAll(CLK := xCmdReadAll);
IF rtReadAll.Q THEN
    RequestReadAll();
END_IF
rtReadIdent(CLK := xCmdReadIdent);
IF rtReadIdent.Q THEN
    RequestReadIdent();
END_IF
rtWrSP1(CLK := xCmdWriteSP1);
IF rtWrSP1.Q THEN
    RequestWrite(iParam := E_O5D150_Param.SP1, diValue := UINT_TO_DINT(uiSetSP1));
END_IF
rtWrLogic(CLK := xCmdWriteLogic);
IF rtWrLogic.Q THEN
    RequestWrite(iParam := E_O5D150_Param.CFG_LOGIC, diValue := USINT_TO_DINT(usiSetLogic));
END_IF
rtWrLaser(CLK := xCmdWriteLaser);
IF rtWrLaser.Q THEN
    RequestWrite(iParam := E_O5D150_Param.LASER, diValue := USINT_TO_DINT(usiSetLaser));
END_IF
rtWrDisplay(CLK := xCmdWriteDisplay);
IF rtWrDisplay.Q THEN
    RequestWrite(iParam := E_O5D150_Param.DISPLAY, diValue := USINT_TO_DINT(usiSetDisplay));
END_IF

// ---------- 3. Align: đọc chu kỳ chậm chỉ khi đang căn chỉnh, tránh chiếm kênh ISDU ----------
tonAlign(IN := xAlignMode AND xPdValid AND NOT tonAlign.Q, PT := tAlignPoll);
IF tonAlign.Q THEN
    RequestRead(E_O5D150_Param.ALIGN);
END_IF

// ---------- 4. Test Event qua System Command (index 2) ----------
rtEvt1On(CLK := xCmdTestEvt1On);
IF rtEvt1On.Q THEN
    QueueSysCmd(GVL_O5D150_Def.usiSC_TEST_EVT1_ON);
END_IF
rtEvt1Off(CLK := xCmdTestEvt1Off);
IF rtEvt1Off.Q THEN
    QueueSysCmd(GVL_O5D150_Def.usiSC_TEST_EVT1_OFF);
END_IF
rtEvt2On(CLK := xCmdTestEvt2On);
IF rtEvt2On.Q THEN
    QueueSysCmd(GVL_O5D150_Def.usiSC_TEST_EVT2_ON);
END_IF
rtEvt2Off(CLK := xCmdTestEvt2Off);
IF rtEvt2Off.Q THEN
    QueueSysCmd(GVL_O5D150_Def.usiSC_TEST_EVT2_OFF);
END_IF
IF usiPendSysCmd <> 0 AND NOT xPendCustom THEN
    abCmd[0] := usiPendSysCmd;
    IF RequestCustom(eService := E_IolService.WRITE, uiIndex := GVL_O5D150_Def.uiIDX_SYS_CMD,
                     usiSubindex := 0, pData := ADR(abCmd), uiLen := 1) THEN
        usiPendSysCmd := 0;
    ELSIF NOT xWriteEnable THEN
        usiPendSysCmd := 0;                     // Maintenance bị tắt giữa chừng: bỏ lệnh
    END_IF
END_IF

// ---------- 5. Danh sách event (index 37). Kênh chính thức là PROFINET diagnosis/alarm của AL1100 (TODO) ----------
IF rtPdValid.Q THEN
    xEvtListNotSupported := FALSE;              // device mới cắm vào: thử lại
END_IF
rtReadEvt(CLK := xCmdReadEvents);
IF rtReadEvt.Q THEN
    xEvtListNotSupported := FALSE;
    xPendEvtRead := TRUE;
END_IF
tonEvt(IN := xPdValid AND NOT xEvtListNotSupported AND NOT tonEvt.Q, PT := tEvtPoll);
IF tonEvt.Q THEN
    xPendEvtRead := TRUE;
END_IF
IF xPendEvtRead AND NOT xPendCustom AND usiPendSysCmd = 0 THEN
    IF RequestCustom(eService := E_IolService.READ, uiIndex := GVL_O5D150_Def.uiIDX_EVT_LIST,
                     usiSubindex := 0, pData := 0, uiLen := 0) THEN
        xPendEvtRead := FALSE;
    END_IF
END_IF

// PDin 16 bit big-endian: Distance 12 bit từ bit 4 [cm], OUT1 bit 0 (layout trong GVL_O5D150_Def.stPdLayout)
METHOD PROTECTED DecodePdIn
VAR
    wRaw   : WORD;
    uiDist : UINT;
END_VAR

(*---IMPL---*)
wRaw := SHL(BYTE_TO_WORD(abPdIn[0]), 8) OR BYTE_TO_WORD(abPdIn[1]);
stPd.wRaw     := wRaw;
stPd.xPdValid := xPdValid;
IF xPdValid THEN
    uiDist := WORD_TO_UINT(SHR(wRaw, GVL_O5D150_Def.stPdLayout.usiDistBitOffset) AND GVL_O5D150_Def.stPdLayout.wDistMask);
    stPd.uiDistance_cm := uiDist;
    stPd.rDistance_m   := UINT_TO_REAL(uiDist) * GVL_O5D150_Def.stPdLayout.rGradient;
    stPd.xOut1         := (SHR(wRaw, GVL_O5D150_Def.stPdLayout.usiOut1Bit) AND WORD#1) <> 0;
    stPd.xOutOfRange   := uiDist < GVL_O5D150_Def.stPdLayout.uiDistMin OR uiDist > GVL_O5D150_Def.stPdLayout.uiDistMax;
ELSE
    // PD không hợp lệ: khoảng cách giữ giá trị cũ để HMI không nhảy về 0, OUT1 về FALSE (fail-safe)
    stPd.xOut1 := FALSE;
END_IF

// Xếp 1 System Command chờ gửi; bị khoá khi chưa bật Maintenance
METHOD PROTECTED QueueSysCmd
VAR_INPUT
    usiCmd : USINT;
END_VAR

(*---IMPL---*)
IF NOT xWriteEnable THEN
    SetLocalErr(E_IolErrSource.WRITE_LOCKED);
ELSE
    usiPendSysCmd := usiCmd;
END_IF

// Giải mã Detailed Device Status (index 37): mỗi entry 3 byte = EventQualifier + EventCode (big-endian),
// entry 0/0 = trống. Đánh dấu cờ theo bảng GVL_O5D150_Def.aEvtDef.
METHOD PROTECTED DecodeEvents
VAR_INPUT
    uiLen : UINT;
END_VAR
VAR
    k      : INT;
    j      : INT;
    wCode  : WORD;
    xFound : BOOL;
END_VAR

(*---IMPL---*)
FOR j := 0 TO GVL_O5D150_Def.iEVT_COUNT - 1 DO
    axEvtActive[j] := FALSE;
END_FOR
uiEvtCount      := 0;
xEvtErrorActive := FALSE;

FOR k := 0 TO UINT_TO_INT(uiLen / 3) - 1 DO
    wCode := UINT_TO_WORD(F_IolGetU16BE(ADR(abBuf), INT_TO_UINT(k * 3 + 1)));
    IF abBuf[k * 3] <> 0 OR wCode <> 0 THEN
        uiEvtCount := uiEvtCount + 1;
        xFound := FALSE;
        FOR j := 0 TO GVL_O5D150_Def.iEVT_COUNT - 1 DO
            IF GVL_O5D150_Def.aEvtDef[j].wCode = wCode THEN
                axEvtActive[j] := TRUE;
                xFound := TRUE;
                IF GVL_O5D150_Def.aEvtDef[j].eType = E_IolEvtType.ERROR THEN
                    xEvtErrorActive := TRUE;
                END_IF
            END_IF
        END_FOR
        IF NOT xFound THEN
            wUnknownEvt := wCode;
        END_IF
    END_IF
END_FOR
xEvtListValid := TRUE;

(*---IMPL---*)
ParamCount := GVL_O5D150_Def.iPARAM_COUNT;

METHOD ParamCount : INT

METHOD GetParamDef : ST_IolParamDef
VAR_INPUT
    iParam : INT;
END_VAR
VAR
    stEmpty : ST_IolParamDef;
END_VAR

(*---IMPL---*)
IF iParam >= 0 AND iParam < GVL_O5D150_Def.iPARAM_COUNT THEN
    GetParamDef := GVL_O5D150_Def.aParamDef[iParam];
ELSE
    GetParamDef := stEmpty;
END_IF

METHOD GetValPtr : POINTER TO ST_IolParamVal
VAR_INPUT
    iParam : INT;
END_VAR

(*---IMPL---*)
IF iParam >= 0 AND iParam < GVL_O5D150_Def.iPARAM_COUNT THEN
    GetValPtr := ADR(aVal[iParam]);
ELSE
    GetValPtr := 0;
END_IF

// Limit (index 64) là record 4 byte: min UINT16 | max UINT16 -> tách ra
METHOD OnParamDone
VAR_INPUT
    iParam : INT;
    xErr   : BOOL;
END_VAR
VAR
    dwRaw : DWORD;
END_VAR

(*---IMPL---*)
IF iParam = E_O5D150_Param.LIMITS AND NOT xErr THEN
    dwRaw := DINT_TO_DWORD(aVal[E_O5D150_Param.LIMITS].diRaw);
    uiLimitMin_cm := DWORD_TO_UINT(SHR(dwRaw, 16));
    uiLimitMax_cm := DWORD_TO_UINT(dwRaw AND 16#FFFF);
END_IF

// Kết quả ISDU tự do: index 37 (event list) và index 2 (System Command)
METHOD OnCustomDone : BOOL
VAR_INPUT
    uiIndex  : UINT;
    eService : E_IolService;
    xErr     : BOOL;
    uiDevErr : UINT;
    uiLen    : UINT;
END_VAR

(*---IMPL---*)
OnCustomDone := FALSE;
IF uiIndex = GVL_O5D150_Def.uiIDX_EVT_LIST AND eService = E_IolService.READ THEN
    IF xErr THEN
        xEvtListValid := FALSE;
        IF uiDevErr = GVL_IolConst.uiERR_IDX_NA THEN
            // IODD không khai báo index 37: ghi nhận 1 lần, ngừng đọc chu kỳ, không đẩy lỗi lên HMI
            xEvtListNotSupported := TRUE;
            OnCustomDone := TRUE;
        END_IF
    ELSE
        DecodeEvents(uiLen);
    END_IF
ELSIF uiIndex = GVL_O5D150_Def.uiIDX_SYS_CMD AND NOT xErr THEN
    xPendEvtRead := TRUE;          // cập nhật danh sách event ngay sau Test Event
END_IF

(* ---- FB_IolCall.st ---- *)
// Client IO-Link Call kiểu PLCopen: sườn lên xExecute -> xBusy -> xDone/xError (giữ tới khi xExecute = FALSE,
// tối thiểu 1 chu kỳ nếu xExecute đã rớt). Request đi qua hàng đợi FB_IolMaster.
FUNCTION_BLOCK FB_IolCall
VAR_INPUT
    refMaster   : REFERENCE TO FB_IolMaster;
    xExecute    : BOOL;
    usiPort     : USINT;                   // 1..4 (0 = master)
    eService    : E_IolService := E_IolService.READ;
    uiIndex     : UINT;
    usiSubindex : USINT;
    pData       : POINTER TO BYTE;         // WRITE: dữ liệu ghi; READ: buffer nhận
    uiDataLen   : UINT;                    // WRITE: số byte ghi; READ: kích thước buffer
END_VAR
VAR_OUTPUT
    xDone          : BOOL;
    xBusy          : BOOL;
    xError         : BOOL;
    uiLenRead      : UINT;
    eErrSource     : E_IolErrSource;
    dwPnioStatus   : DWORD;
    uiIolMasterErr : UINT;
    uiIolDevErr    : UINT;
    wsErrText      : WSTRING(80);
END_VAR
VAR
    rtExec  : R_TRIG;
    eStep   : E_IolCallStep;
    hHandle : USINT;                       // handle đăng ký với master (1 lần)
    stReq   : ST_IolRequest;
    stRes   : ST_IolResult;
    tonWait : TON;                         // timeout phía client, bao cả thời gian chờ hàng đợi
    i       : INT;
    n       : UINT;
END_VAR

(*---IMPL---*)
rtExec(CLK := xExecute);

CASE eStep OF
    E_IolCallStep.IDLE:
        xDone  := FALSE;
        xError := FALSE;
        xBusy  := FALSE;
        tonWait(IN := FALSE);
        IF rtExec.Q THEN
            uiLenRead := 0;
            eErrSource := E_IolErrSource.NONE;
            dwPnioStatus := 0;
            uiIolMasterErr := 0;
            uiIolDevErr := 0;
            wsErrText := "";
            // kiểm tham số trước khi gửi
            IF NOT __ISVALIDREF(refMaster) OR usiPort > 4 OR pData = 0
               OR uiDataLen > GVL_IolConst.uiMAX_DATA
               OR (eService = E_IolService.WRITE AND uiDataLen = 0) THEN
                SetError(E_IolErrSource.PARAM);
            ELSE
                IF hHandle = 0 THEN
                    hHandle := refMaster.Register();
                END_IF
                stReq.usiPort     := usiPort;
                stReq.eService    := eService;
                stReq.uiIndex     := uiIndex;
                stReq.usiSubindex := usiSubindex;
                stReq.uiLen       := 0;
                IF eService = E_IolService.WRITE THEN
                    stReq.uiLen := uiDataLen;
                    FOR i := 0 TO UINT_TO_INT(uiDataLen) - 1 DO
                        stReq.abData[i] := pData[i];
                    END_FOR
                END_IF
                IF hHandle = 0 THEN
                    SetError(E_IolErrSource.LOCK);
                ELSIF refMaster.Submit(hHandle := hHandle, stReq := stReq) THEN
                    xBusy := TRUE;
                    eStep := E_IolCallStep.WAIT;
                ELSE
                    SetError(E_IolErrSource.LOCK);
                END_IF
            END_IF
        END_IF

    E_IolCallStep.WAIT:
        xBusy := TRUE;
        tonWait(IN := TRUE, PT := refMaster.tTimeout * 2);
        IF refMaster.Poll(hHandle := hHandle, stRes := stRes) THEN
            tonWait(IN := FALSE);
            xBusy := FALSE;
            IF stRes.xError THEN
                dwPnioStatus   := stRes.dwPnioStatus;
                uiIolMasterErr := stRes.uiIolMasterErr;
                uiIolDevErr    := stRes.uiIolDevErr;
                SetError(stRes.eErrSource);
            ELSE
                IF eService = E_IolService.READ THEN
                    n := MIN(stRes.uiLen, uiDataLen);
                    FOR i := 0 TO UINT_TO_INT(n) - 1 DO
                        pData[i] := stRes.abData[i];
                    END_FOR
                    uiLenRead := n;
                END_IF
                xDone := TRUE;
                eStep := E_IolCallStep.DONE;
            END_IF
        ELSIF tonWait.Q THEN
            tonWait(IN := FALSE);
            refMaster.Cancel(hHandle := hHandle);
            xBusy := FALSE;
            SetError(E_IolErrSource.TIMEOUT);
        END_IF

    E_IolCallStep.DONE:
        xBusy := FALSE;
        xDone := TRUE;
        IF NOT xExecute THEN
            eStep := E_IolCallStep.IDLE;      // chu kỳ sau IDLE mới xoá xDone
        END_IF

    E_IolCallStep.ERR:
        xBusy  := FALSE;
        xError := TRUE;
        IF NOT xExecute THEN
            eStep := E_IolCallStep.IDLE;
        END_IF
END_CASE

// Chuyển sang ERR, ghi nguồn lỗi + chuỗi hiển thị
METHOD PRIVATE SetError
VAR_INPUT
    eSrc : E_IolErrSource;
END_VAR

(*---IMPL---*)
eErrSource := eSrc;
wsErrText  := F_IolErrText(eSrc, uiIolMasterErr, uiIolDevErr, dwPnioStatus);
xBusy  := FALSE;
xDone  := FALSE;
xError := TRUE;
eStep  := E_IolCallStep.ERR;

(* ---- FB_IolDevBase.st ---- *)
// Lớp cơ sở cho mọi device IO-Link: giải mã PQI, trình tự đọc/ghi tham số theo bảng IODD của lớp con,
// đọc Ident 16..24, kênh ISDU tự do cho lớp con. Lớp con override: ParamCount, GetParamDef, GetValPtr,
// OnParamDone, OnCustomDone và gọi SUPER^() trong thân.
FUNCTION_BLOCK FB_IolDevBase
VAR_INPUT
    refMaster          : REFERENCE TO FB_IolMaster;
    usiPort            : USINT;
    bPQI               : BYTE;                  // Port Qualifier từ GVL_IO
    xWriteEnable       : BOOL;                  // khoá ghi tham số / System Command (Maintenance)
    xAutoReadOnConnect : BOOL := TRUE;          // tự đọc Ident + ReadAll khi PD chuyển hợp lệ
    xResetErr          : BOOL;                  // sườn lên: xoá lỗi gần nhất
END_VAR
VAR_OUTPUT
    stDiag         : ST_IolPortDiag;
    xPdValid       : BOOL;                      // PQ AND DA
    xBusy          : BOOL;                      // đang chạy hoặc còn việc chờ
    xLastError     : BOOL;                      // lỗi gần nhất, giữ tới xResetErr
    eLastErrSrc    : E_IolErrSource;
    uiLastDevErr   : UINT;
    wsLastErr      : WSTRING(80);
    stIdent        : ST_IolIdent;
    udiJobCount    : UDINT;
    udiJobErrCount : UDINT;
END_VAR
VAR
    fbCall      : FB_IolCall;                   // instance riêng mỗi device
    eSeq        : E_IolDevSeq;
    eJob        : E_IolDevJob;
    iJobParam   : INT;
    uiJobIndex  : UINT;
    usiJobSub   : USINT;
    eJobService : E_IolService := E_IolService.READ;
    uiJobLen    : UINT;
    xCallExec   : BOOL;
    abBuf       : ARRAY[0..GVL_IolConst.uiMAX_DATA - 1] OF BYTE;   // dữ liệu ghi / nhận của việc đang chạy
    axPendRead  : ARRAY[0..GVL_IolConst.iMAX_PARAM - 1] OF BOOL;
    axPendWrite : ARRAY[0..GVL_IolConst.iMAX_PARAM - 1] OF BOOL;
    wPendIdent  : WORD;                         // bit n = cần đọc index 16 + n
    xPendCustom : BOOL;
    stCustom    : ST_IolRequest;
    rtPdValid   : R_TRIG;
    rtResetErr  : R_TRIG;
END_VAR

(*---IMPL---*)
// ---------- 1. Port Qualifier (bit theo GSDML AL1100) ----------
stDiag.bPQI := bPQI;
stDiag.xDI4 := bPQI.0;
stDiag.xDI2 := bPQI.1;
stDiag.xNP  := bPQI.2;
stDiag.xSV  := bPQI.3;
stDiag.xDA  := bPQI.4;
stDiag.xDC  := bPQI.5;
stDiag.xDE  := bPQI.6;
stDiag.xPQ  := bPQI.7;
xPdValid := stDiag.xPQ AND stDiag.xDA;

rtPdValid(CLK := xPdValid);
IF rtPdValid.Q AND xAutoReadOnConnect THEN
    RequestReadIdent();
    RequestReadAll();
END_IF

rtResetErr(CLK := xResetErr);
IF rtResetErr.Q THEN
    xLastError   := FALSE;
    eLastErrSrc  := E_IolErrSource.NONE;
    uiLastDevErr := 0;
    wsLastErr    := "";
END_IF

// ---------- 2. Port không có thiết bị: huỷ việc chờ ngay, không đợi timeout ----------
IF NOT stDiag.xDA AND eSeq = E_IolDevSeq.IDLE AND HasPending() THEN
    DropAll();
END_IF

// ---------- 3. Client IOL_CALL: gọi đúng 1 lần mỗi chu kỳ ----------
IF __ISVALIDREF(refMaster) THEN
    fbCall.refMaster REF= refMaster;
END_IF
IF eJobService = E_IolService.WRITE THEN
    fbCall(xExecute := xCallExec, usiPort := usiPort, eService := eJobService, uiIndex := uiJobIndex,
           usiSubindex := usiJobSub, pData := ADR(abBuf), uiDataLen := uiJobLen);
ELSE
    fbCall(xExecute := xCallExec, usiPort := usiPort, eService := eJobService, uiIndex := uiJobIndex,
           usiSubindex := usiJobSub, pData := ADR(abBuf), uiDataLen := GVL_IolConst.uiMAX_DATA);
END_IF

// ---------- 4. Trình tự việc ----------
CASE eSeq OF
    E_IolDevSeq.IDLE:
        xCallExec := FALSE;
        IF SelectJob() THEN
            xCallExec := TRUE;
            eSeq := E_IolDevSeq.RUN;
        END_IF

    E_IolDevSeq.RUN:
        IF fbCall.xDone OR fbCall.xError THEN
            xCallExec := FALSE;
            JobFinished(xErr := fbCall.xError);
            eSeq := E_IolDevSeq.RELEASE;
        END_IF

    E_IolDevSeq.RELEASE:
        // chờ FB_IolCall về IDLE để sườn Execute kế tiếp chắc chắn được nhận
        IF NOT fbCall.xDone AND NOT fbCall.xError AND NOT fbCall.xBusy THEN
            eJob := E_IolDevJob.NONE;
            eSeq := E_IolDevSeq.IDLE;
        END_IF
END_CASE

xBusy := (eSeq <> E_IolDevSeq.IDLE) OR HasPending();

(*---IMPL---*)
ParamCount := 0;

// Số tham số trong bảng IODD của device - lớp con override
METHOD ParamCount : INT

// Định nghĩa tham số thứ iParam - lớp con override
METHOD GetParamDef : ST_IolParamDef
VAR_INPUT
    iParam : INT;
END_VAR
VAR
    stEmpty : ST_IolParamDef;
END_VAR

(*---IMPL---*)
GetParamDef := stEmpty;

// Con trỏ tới giá trị runtime của tham số iParam (mảng nằm ở lớp con); 0 = không có
METHOD GetValPtr : POINTER TO ST_IolParamVal
VAR_INPUT
    iParam : INT;
END_VAR

(*---IMPL---*)
GetValPtr := 0;

// Hook sau khi đọc xong 1 tham số (lớp con tách record nhiều trường...)
METHOD OnParamDone
VAR_INPUT
    iParam : INT;
    xErr   : BOOL;
END_VAR

(*---IMPL---*)
;

// Hook khi việc ISDU tự do kết thúc; dữ liệu đọc nằm trong abBuf[0..uiLen-1].
// Trả TRUE để KHÔNG đẩy lỗi lên wsLastErr (lớp con tự xử lý, vd index không hỗ trợ).
METHOD OnCustomDone : BOOL
VAR_INPUT
    uiIndex  : UINT;
    eService : E_IolService;
    xErr     : BOOL;
    uiDevErr : UINT;
    uiLen    : UINT;
END_VAR

(*---IMPL---*)
OnCustomDone := FALSE;

// Đánh dấu đọc mọi tham số có xInReadAll và không phải write-only
METHOD RequestReadAll
VAR
    i     : INT;
    stDef : ST_IolParamDef;
END_VAR

(*---IMPL---*)
FOR i := 0 TO MIN(THIS^.ParamCount(), GVL_IolConst.iMAX_PARAM) - 1 DO
    stDef := THIS^.GetParamDef(i);
    IF stDef.xInReadAll AND stDef.eAccess <> E_IolAccess.WO THEN
        axPendRead[i] := TRUE;
    END_IF
END_FOR

(*---IMPL---*)
wPendIdent := 16#01FF;

// Đánh dấu đọc Ident index 16..24
METHOD RequestReadIdent

// Đánh dấu đọc 1 tham số; FALSE nếu iParam sai hoặc tham số write-only
METHOD RequestRead : BOOL
VAR_INPUT
    iParam : INT;
END_VAR
VAR
    stDef : ST_IolParamDef;
END_VAR

(*---IMPL---*)
RequestRead := FALSE;
IF iParam < 0 OR iParam >= MIN(THIS^.ParamCount(), GVL_IolConst.iMAX_PARAM) THEN
    RETURN;
END_IF
stDef := THIS^.GetParamDef(iParam);
IF stDef.eAccess = E_IolAccess.WO THEN
    RETURN;
END_IF
axPendRead[iParam] := TRUE;
RequestRead := TRUE;

// Yêu cầu ghi 1 tham số. Chặn trước khi gửi: khoá ghi (xWriteEnable), tham số read-only, ngoài dải IODD.
// Ghi xong tự đọc lại để xác nhận.
METHOD RequestWrite : BOOL
VAR_INPUT
    iParam  : INT;
    diValue : DINT;
END_VAR
VAR
    stDef : ST_IolParamDef;
    pVal  : POINTER TO ST_IolParamVal;
END_VAR

(*---IMPL---*)
RequestWrite := FALSE;
IF iParam < 0 OR iParam >= MIN(THIS^.ParamCount(), GVL_IolConst.iMAX_PARAM) THEN
    SetLocalErr(E_IolErrSource.PARAM);
    RETURN;
END_IF
stDef := THIS^.GetParamDef(iParam);
pVal  := THIS^.GetValPtr(iParam);
IF pVal = 0 OR stDef.eAccess = E_IolAccess.RO THEN
    SetLocalErr(E_IolErrSource.PARAM);
    RETURN;
END_IF
IF NOT xWriteEnable THEN
    SetLocalErr(E_IolErrSource.WRITE_LOCKED);
    RETURN;
END_IF
IF diValue < stDef.diMin OR diValue > stDef.diMax THEN
    pVal^.uiErr := 16#FF00 OR INT_TO_UINT(E_IolErrSource.RANGE);
    SetLocalErr(E_IolErrSource.RANGE);
    RETURN;
END_IF
pVal^.diSet  := diValue;
pVal^.xDirty := TRUE;
axPendWrite[iParam] := TRUE;
RequestWrite := TRUE;

// ISDU tự do (System Command, event list...). 1 việc chờ tại 1 thời điểm; FALSE nếu đang có việc chờ,
// ghi bị khoá hoặc độ dài sai. Kết quả báo qua OnCustomDone.
METHOD RequestCustom : BOOL
VAR_INPUT
    eService    : E_IolService;
    uiIndex     : UINT;
    usiSubindex : USINT;
    pData       : POINTER TO BYTE;     // chỉ dùng khi WRITE
    uiLen       : UINT;                // số byte ghi (READ bỏ qua)
END_VAR
VAR
    i : INT;
END_VAR

(*---IMPL---*)
RequestCustom := FALSE;
IF xPendCustom THEN
    RETURN;
END_IF
IF eService = E_IolService.WRITE THEN
    IF NOT xWriteEnable THEN
        SetLocalErr(E_IolErrSource.WRITE_LOCKED);
        RETURN;
    END_IF
    IF pData = 0 OR uiLen = 0 OR uiLen > GVL_IolConst.uiMAX_DATA THEN
        SetLocalErr(E_IolErrSource.PARAM);
        RETURN;
    END_IF
    FOR i := 0 TO UINT_TO_INT(uiLen) - 1 DO
        stCustom.abData[i] := pData[i];
    END_FOR
    stCustom.uiLen := uiLen;
ELSE
    stCustom.uiLen := 0;
END_IF
stCustom.usiPort     := usiPort;
stCustom.eService    := eService;
stCustom.uiIndex     := uiIndex;
stCustom.usiSubindex := usiSubindex;
xPendCustom := TRUE;
RequestCustom := TRUE;

// Ghi lỗi phát sinh trong PLC (không qua ISDU) vào lỗi gần nhất
METHOD PROTECTED SetLocalErr
VAR_INPUT
    eSrc : E_IolErrSource;
END_VAR

(*---IMPL---*)
xLastError   := TRUE;
eLastErrSrc  := eSrc;
uiLastDevErr := 0;
wsLastErr    := F_IolErrText(eSrc, 0, 0, 0);

(*---IMPL---*)
xLastError   := TRUE;
eLastErrSrc  := fbCall.eErrSource;
uiLastDevErr := fbCall.uiIolDevErr;
wsLastErr    := fbCall.wsErrText;

// Chép lỗi của lần gọi ISDU vừa xong vào lỗi gần nhất
METHOD PROTECTED ReportErr

(*---IMPL---*)
IF fbCall.uiIolDevErr <> 0 THEN
    ErrCode := fbCall.uiIolDevErr;
ELSE
    ErrCode := 16#FF00 OR INT_TO_UINT(fbCall.eErrSource);
END_IF

// Mã lỗi lưu vào ST_IolParamVal.uiErr: lỗi device 0x80xx, còn lại 0xFF00 + E_IolErrSource
METHOD PROTECTED ErrCode : UINT

// Còn việc ISDU nào đang chờ không
METHOD PROTECTED HasPending : BOOL
VAR
    i : INT;
END_VAR

(*---IMPL---*)
HasPending := xPendCustom OR (wPendIdent <> 0);
FOR i := 0 TO GVL_IolConst.iMAX_PARAM - 1 DO
    IF axPendRead[i] OR axPendWrite[i] THEN
        HasPending := TRUE;
        RETURN;
    END_IF
END_FOR

// Huỷ mọi việc chờ khi port không có thiết bị, báo NO_DEVICE thay vì để từng request timeout
METHOD PROTECTED DropAll
VAR
    i : INT;
END_VAR

(*---IMPL---*)
FOR i := 0 TO GVL_IolConst.iMAX_PARAM - 1 DO
    axPendRead[i]  := FALSE;
    axPendWrite[i] := FALSE;
END_FOR
wPendIdent := 0;
IF xPendCustom THEN
    xPendCustom := FALSE;
    THIS^.OnCustomDone(uiIndex := stCustom.uiIndex, eService := stCustom.eService, xErr := TRUE, uiDevErr := 0, uiLen := 0);
END_IF
SetLocalErr(E_IolErrSource.NO_DEVICE);

// Chọn việc tiếp theo theo ưu tiên: tự do (System Command / event) > ghi > đọc tham số > Ident
METHOD PROTECTED SelectJob : BOOL
VAR
    i     : INT;
    iN    : INT;
    stDef : ST_IolParamDef;
END_VAR

(*---IMPL---*)
SelectJob := FALSE;
IF NOT stDiag.xDA THEN
    RETURN;
END_IF
iN := MIN(THIS^.ParamCount(), GVL_IolConst.iMAX_PARAM);

// --- 1. ISDU tự do ---
IF xPendCustom THEN
    xPendCustom := FALSE;
    eJob        := E_IolDevJob.CUSTOM;
    iJobParam   := -1;
    uiJobIndex  := stCustom.uiIndex;
    usiJobSub   := stCustom.usiSubindex;
    eJobService := stCustom.eService;
    uiJobLen    := stCustom.uiLen;
    FOR i := 0 TO UINT_TO_INT(stCustom.uiLen) - 1 DO
        abBuf[i] := stCustom.abData[i];
    END_FOR
    SelectJob := TRUE;
    RETURN;
END_IF

// --- 2. Ghi tham số ---
FOR i := 0 TO iN - 1 DO
    IF axPendWrite[i] THEN
        axPendWrite[i] := FALSE;
        IF PrepareWrite(i) THEN
            eJob := E_IolDevJob.PARAM_WR;
            SelectJob := TRUE;
            RETURN;
        END_IF
    END_IF
END_FOR

// --- 3. Đọc tham số ---
FOR i := 0 TO iN - 1 DO
    IF axPendRead[i] THEN
        axPendRead[i] := FALSE;
        stDef := THIS^.GetParamDef(i);
        eJob        := E_IolDevJob.PARAM_RD;
        iJobParam   := i;
        uiJobIndex  := stDef.uiIndex;
        usiJobSub   := stDef.usiSubindex;
        eJobService := E_IolService.READ;
        uiJobLen    := 0;
        SelectJob := TRUE;
        RETURN;
    END_IF
END_FOR

// --- 4. Ident 16..24 ---
IF wPendIdent <> 0 THEN
    FOR i := 0 TO 8 DO
        IF (SHR(wPendIdent, i) AND WORD#1) <> 0 THEN
            wPendIdent  := wPendIdent AND NOT SHL(WORD#1, i);
            eJob        := E_IolDevJob.IDENT;
            iJobParam   := -1;
            uiJobIndex  := 16 + INT_TO_UINT(i);
            usiJobSub   := 0;
            eJobService := E_IolService.READ;
            uiJobLen    := 0;
            SelectJob := TRUE;
            RETURN;
        END_IF
    END_FOR
    wPendIdent := 0;
END_IF

// Mã hoá diSet của tham số iParam thành byte big-endian trong abBuf; FALSE nếu kiểu không hỗ trợ ghi qua bảng
METHOD PROTECTED PrepareWrite : BOOL
VAR_INPUT
    iParam : INT;
END_VAR
VAR
    stDef : ST_IolParamDef;
    pVal  : POINTER TO ST_IolParamVal;
END_VAR

(*---IMPL---*)
PrepareWrite := FALSE;
stDef := THIS^.GetParamDef(iParam);
pVal  := THIS^.GetValPtr(iParam);
IF pVal = 0 THEN
    RETURN;
END_IF
iJobParam   := iParam;
uiJobIndex  := stDef.uiIndex;
usiJobSub   := stDef.usiSubindex;
eJobService := E_IolService.WRITE;
CASE stDef.eType OF
    E_IolDataType.U8, E_IolDataType.I8:
        abBuf[0] := DINT_TO_BYTE(pVal^.diSet);
        uiJobLen := 1;
    E_IolDataType.U16, E_IolDataType.I16:
        F_IolSetU16BE(ADR(abBuf), 0, DINT_TO_UINT(pVal^.diSet));
        uiJobLen := 2;
    E_IolDataType.U32, E_IolDataType.I32:
        F_IolSetU32BE(ADR(abBuf), 0, DINT_TO_DWORD(pVal^.diSet));
        uiJobLen := 4;
ELSE
    pVal^.xDirty := FALSE;
    RETURN;
END_CASE
PrepareWrite := TRUE;

// Giải mã abBuf (big-endian) thành diRaw của tham số iParam
METHOD PROTECTED DecodeParam
VAR_INPUT
    iParam : INT;
    uiLen  : UINT;
END_VAR
VAR
    stDef  : ST_IolParamDef;
    pVal   : POINTER TO ST_IolParamVal;
    uiNeed : UINT;
END_VAR

(*---IMPL---*)
stDef := THIS^.GetParamDef(iParam);
pVal  := THIS^.GetValPtr(iParam);
IF pVal = 0 THEN
    RETURN;
END_IF
CASE stDef.eType OF
    E_IolDataType.U8, E_IolDataType.I8:   uiNeed := 1;
    E_IolDataType.U16, E_IolDataType.I16: uiNeed := 2;
ELSE
    uiNeed := 4;
END_CASE
IF uiLen < uiNeed THEN
    pVal^.xValid := FALSE;
    pVal^.uiErr  := 16#FF00 OR INT_TO_UINT(E_IolErrSource.FRAME);
    RETURN;
END_IF
CASE stDef.eType OF
    E_IolDataType.U8:  pVal^.diRaw := BYTE_TO_DINT(abBuf[0]);
    E_IolDataType.I8:  pVal^.diRaw := SINT_TO_DINT(BYTE_TO_SINT(abBuf[0]));
    E_IolDataType.U16: pVal^.diRaw := UINT_TO_DINT(F_IolGetU16BE(ADR(abBuf), 0));
    E_IolDataType.I16: pVal^.diRaw := INT_TO_DINT(UINT_TO_INT(F_IolGetU16BE(ADR(abBuf), 0)));
ELSE
    pVal^.diRaw := DWORD_TO_DINT(F_IolGetU32BE(ADR(abBuf), 0));   // U32/I32/OCTET 4 byte đầu
END_CASE
pVal^.xValid := TRUE;
pVal^.uiErr  := 0;

// Lưu chuỗi Ident vừa đọc (abBuf) vào stIdent
METHOD PROTECTED StoreIdent
VAR_INPUT
    uiIndex : UINT;
    uiLen   : UINT;
END_VAR
VAR
    sVal : STRING(64);
END_VAR

(*---IMPL---*)
sVal := F_IolBytesToStr(ADR(abBuf), uiLen);
CASE uiIndex OF
    16: stIdent.sVendorName  := sVal;
    17: stIdent.sVendorText  := sVal;
    18: stIdent.sProductName := sVal;
    19: stIdent.sProductId   := sVal;
    20: stIdent.sProductText := sVal;
    21: stIdent.sSerialNo    := sVal;
    22: stIdent.sHwRev       := sVal;
    23: stIdent.sFwRev       := sVal;
    24: stIdent.sAppTag      := sVal;
END_CASE

// Xử lý kết quả của việc vừa xong
METHOD PROTECTED JobFinished
VAR_INPUT
    xErr : BOOL;
END_VAR
VAR
    pVal : POINTER TO ST_IolParamVal;
END_VAR

(*---IMPL---*)
udiJobCount := udiJobCount + 1;
IF xErr THEN
    udiJobErrCount := udiJobErrCount + 1;
END_IF

CASE eJob OF
    E_IolDevJob.PARAM_RD:
        pVal := THIS^.GetValPtr(iJobParam);
        IF pVal <> 0 THEN
            IF xErr THEN
                pVal^.xValid := FALSE;
                pVal^.uiErr  := ErrCode();
            ELSE
                DecodeParam(iJobParam, fbCall.uiLenRead);
            END_IF
        END_IF
        IF xErr THEN
            ReportErr();
        END_IF
        THIS^.OnParamDone(iParam := iJobParam, xErr := xErr);

    E_IolDevJob.PARAM_WR:
        pVal := THIS^.GetValPtr(iJobParam);
        IF pVal <> 0 THEN
            pVal^.xDirty := FALSE;
            IF xErr THEN
                pVal^.uiErr := ErrCode();
            ELSE
                pVal^.uiErr := 0;
                axPendRead[iJobParam] := TRUE;     // đọc lại để xác nhận giá trị device đã nhận
            END_IF
        END_IF
        IF xErr THEN
            ReportErr();
        END_IF

    E_IolDevJob.IDENT:
        // index Ident là tuỳ chọn theo device: lỗi thì bỏ qua, giữ chuỗi rỗng
        IF NOT xErr THEN
            StoreIdent(uiJobIndex, fbCall.uiLenRead);
        END_IF

    E_IolDevJob.CUSTOM:
        IF NOT THIS^.OnCustomDone(uiIndex := uiJobIndex, eService := eJobService, xErr := xErr,
                                  uiDevErr := fbCall.uiIolDevErr, uiLen := fbCall.uiLenRead) AND xErr THEN
            ReportErr();
        END_IF
END_CASE

(* ---- FB_IolMaster.st ---- *)
// 1 instance cho mỗi IO-Link master (AL1100). Khoá + hàng đợi FIFO: tại 1 thời điểm chỉ 1 IOL_CALL
// chạy trên record CAP, các client (FB_IolCall) lần lượt theo thứ tự Submit -> công bằng giữa các device.
FUNCTION_BLOCK FB_IolMaster
VAR_INPUT
    itfRec   : ITF_IolRecordAccess;                // transport thật (FB_PnRecordAccess) hoặc mock
    xEnable  : BOOL := TRUE;                       // FALSE: không lấy request mới từ hàng đợi
    dwId     : DWORD;                              // ID submodule CAP (CommFB.SUBSLOT_ID), mock bỏ qua
    tTimeout : TIME := GVL_IolConst.tCALL_TIMEOUT;
    xReset   : BOOL;                               // xoá hàng đợi, thoát STUCK
END_VAR
VAR_OUTPUT
    eState          : E_IolCallState;
    xBusy           : BOOL;
    usiActiveClient : USINT;                       // handle đang chạy, 0 = rảnh
    uiQueueCount    : UINT;
    udiCallCount    : UDINT;                       // số lần gọi OK
    udiErrCount     : UDINT;                       // số lần gọi lỗi
    xNoTransport    : BOOL;                        // itfRec chưa gán
END_VAR
VAR
    aQueue     : ARRAY[0..GVL_IolConst.iQUEUE_SIZE - 1] OF USINT;   // FIFO handle
    iHead      : INT;
    iCount     : INT;
    aReq       : ARRAY[1..GVL_IolConst.iQUEUE_SIZE] OF ST_IolRequest;
    aRes       : ARRAY[1..GVL_IolConst.iQUEUE_SIZE] OF ST_IolResult;
    axPending  : ARRAY[1..GVL_IolConst.iQUEUE_SIZE] OF BOOL;        // đã Submit, chưa có kết quả
    axResReady : ARRAY[1..GVL_IolConst.iQUEUE_SIZE] OF BOOL;        // kết quả chờ client Poll
    axCancel   : ARRAY[1..GVL_IolConst.iQUEUE_SIZE] OF BOOL;        // client đã bỏ, huỷ kết quả
    usiHandles : USINT;                                             // số client đã Register
    abTx       : ARRAY[0..GVL_IolConst.uiMAX_REC - 1] OF BYTE;      // khung gửi (Watch khi test)
    abRx       : ARRAY[0..GVL_IolConst.uiMAX_REC - 1] OF BYTE;      // khung nhận
    uiTxLen    : UINT;
    uiRxLen    : UINT;
    xWrReq     : BOOL;          // REQ cho chu kỳ sau (state machine quyết định)
    xRdReq     : BOOL;
    xWrDone    : BOOL;
    xWrBusy    : BOOL;
    xWrErr     : BOOL;
    dwWrStatus : DWORD;
    xRdValid   : BOOL;
    xRdBusy    : BOOL;
    xRdErr     : BOOL;
    dwRdStatus : DWORD;
    iRdLen     : INT;
    tonTimeout : TON;
    tonRetry   : TON;
    tonStuck   : TON;
    iRetry     : INT;
    stCur      : ST_IolResult;  // kết quả request đang chạy
    stEmpty    : ST_IolResult;
    i          : INT;
END_VAR

(*---IMPL---*)
// ---------- 0. Reset: trả lỗi LOCK cho mọi request đang chờ, về IDLE ----------
IF xReset THEN
    xWrReq := FALSE;
    xRdReq := FALSE;
    FOR i := 1 TO GVL_IolConst.iQUEUE_SIZE DO
        IF axPending[i] AND NOT axCancel[i] THEN
            aRes[i] := stEmpty;
            aRes[i].xError := TRUE;
            aRes[i].eErrSource := E_IolErrSource.LOCK;
            axResReady[i] := TRUE;
        END_IF
        axPending[i] := FALSE;
        axCancel[i]  := FALSE;
    END_FOR
    iHead := 0;
    iCount := 0;
    usiActiveClient := 0;
    tonTimeout(IN := FALSE);
    tonRetry(IN := FALSE);
    tonStuck(IN := FALSE);
    eState := E_IolCallState.IDLE;
END_IF

// ---------- 1. Gọi transport đúng 1 lần mỗi chu kỳ, REQ do chu kỳ trước quyết định ----------
xNoTransport := (itfRec = 0);
IF NOT xNoTransport THEN
    itfRec.Write(xReq := xWrReq, dwId := dwId, iIndex := UINT_TO_INT(GVL_IolConst.uiCAP_INDEX),
                 iLen := UINT_TO_INT(uiTxLen), pData := ADR(abTx),
                 xDone => xWrDone, xBusy => xWrBusy, xError => xWrErr, dwStatus => dwWrStatus);
    itfRec.Read(xReq := xRdReq, dwId := dwId, iIndex := UINT_TO_INT(GVL_IolConst.uiCAP_INDEX),
                iMLen := UINT_TO_INT(GVL_IolConst.uiMAX_REC), pData := ADR(abRx),
                xValid => xRdValid, xBusy => xRdBusy, xError => xRdErr, dwStatus => dwRdStatus, iLen => iRdLen);
ELSE
    xWrDone := FALSE; xWrBusy := FALSE; xWrErr := FALSE;
    xRdValid := FALSE; xRdBusy := FALSE; xRdErr := FALSE;
END_IF

// ---------- 2. Timeout tổng của 1 request ----------
tonTimeout(IN := eState = E_IolCallState.WRITE_REQ OR eState = E_IolCallState.RETRY_WR
              OR eState = E_IolCallState.READ_WAIT OR eState = E_IolCallState.READ_REQ,
           PT := tTimeout);
IF tonTimeout.Q THEN
    xWrReq := FALSE;
    xRdReq := FALSE;
    tonStuck(IN := FALSE);
    eState := E_IolCallState.TIMEOUT;
END_IF

// ---------- 3. State machine IOL_CALL ----------
CASE eState OF
    E_IolCallState.IDLE:
        xWrReq := FALSE;
        xRdReq := FALSE;
        IF xEnable AND iCount > 0 THEN
            usiActiveClient := aQueue[iHead];
            iHead  := (iHead + 1) MOD GVL_IolConst.iQUEUE_SIZE;
            iCount := iCount - 1;
            IF axCancel[usiActiveClient] OR NOT axPending[usiActiveClient] THEN
                // client đã bỏ trước khi tới lượt: bỏ qua, không gửi
                axCancel[usiActiveClient]  := FALSE;
                axPending[usiActiveClient] := FALSE;
                usiActiveClient := 0;
            ELSE
                stCur  := stEmpty;
                iRetry := 0;
                BuildFrame();
                IF xNoTransport THEN
                    stCur.eErrSource   := E_IolErrSource.PNIO;
                    stCur.dwPnioStatus := GVL_IolConst.dwSTAT_NO_TRANSPORT;
                    eState := E_IolCallState.ERROR;
                ELSE
                    xWrReq := TRUE;
                    eState := E_IolCallState.WRITE_REQ;
                END_IF
            END_IF
        END_IF

    E_IolCallState.WRITE_REQ:
        IF xWrDone THEN
            xWrReq := FALSE;
            tonRetry(IN := FALSE);
            eState := E_IolCallState.READ_WAIT;
        ELSIF xWrErr THEN
            xWrReq := FALSE;
            IF F_IolIsPnioBusy(dwWrStatus) AND iRetry < GVL_IolConst.iMAX_RETRY THEN
                iRetry := iRetry + 1;
                tonRetry(IN := FALSE);
                eState := E_IolCallState.RETRY_WR;
            ELSE
                stCur.eErrSource   := E_IolErrSource.PNIO;
                stCur.dwPnioStatus := dwWrStatus;
                eState := E_IolCallState.ERROR;
            END_IF
        END_IF

    E_IolCallState.RETRY_WR:
        tonRetry(IN := TRUE, PT := GVL_IolConst.tRETRY_DELAY);
        IF tonRetry.Q THEN
            tonRetry(IN := FALSE);
            xWrReq := TRUE;
            eState := E_IolCallState.WRITE_REQ;
        END_IF

    E_IolCallState.READ_WAIT:
        tonRetry(IN := TRUE, PT := GVL_IolConst.tRETRY_DELAY);
        IF tonRetry.Q THEN
            tonRetry(IN := FALSE);
            xRdReq := TRUE;
            eState := E_IolCallState.READ_REQ;
        END_IF

    E_IolCallState.READ_REQ:
        IF xRdValid THEN
            xRdReq  := FALSE;
            uiRxLen := INT_TO_UINT(MAX(iRdLen, 0));
            IF ParseResponse() THEN
                eState := E_IolCallState.DONE;
            ELSE
                eState := E_IolCallState.ERROR;
            END_IF
        ELSIF xRdErr THEN
            xRdReq := FALSE;
            IF F_IolIsPnioBusy(dwRdStatus) AND iRetry < GVL_IolConst.iMAX_RETRY THEN
                iRetry := iRetry + 1;                 // ISDU chưa xong trên master -> đọc lại sau
                tonRetry(IN := FALSE);
                eState := E_IolCallState.READ_WAIT;
            ELSE
                stCur.eErrSource   := E_IolErrSource.PNIO;
                stCur.dwPnioStatus := dwRdStatus;
                eState := E_IolCallState.ERROR;
            END_IF
        END_IF

    E_IolCallState.DONE:
        Finish(xErr := FALSE);
        eState := E_IolCallState.IDLE;

    E_IolCallState.ERROR:
        Finish(xErr := TRUE);
        eState := E_IolCallState.IDLE;

    E_IolCallState.TIMEOUT:
        // REQ đã hạ; chờ transport hết BUSY rồi mới cho request mới (tránh chồng record)
        xWrReq := FALSE;
        xRdReq := FALSE;
        tonStuck(IN := TRUE, PT := T#1S);
        IF NOT xWrBusy AND NOT xRdBusy THEN
            tonStuck(IN := FALSE);
            stCur.eErrSource := E_IolErrSource.TIMEOUT;
            Finish(xErr := TRUE);
            eState := E_IolCallState.IDLE;
        ELSIF tonStuck.Q THEN
            tonStuck(IN := FALSE);
            stCur.eErrSource := E_IolErrSource.TIMEOUT;
            Finish(xErr := TRUE);
            eState := E_IolCallState.STUCK;
        END_IF

    E_IolCallState.STUCK:
        // chỉ thoát bằng xReset (bước 0)
        xWrReq := FALSE;
        xRdReq := FALSE;
END_CASE

xBusy := (eState <> E_IolCallState.IDLE);
uiQueueCount := INT_TO_UINT(iCount);

// Tạo khung IOL_CALL (abTx, uiTxLen) cho client đang chạy - layout plan mục 4.2
METHOD PRIVATE BuildFrame
VAR
    h : USINT;
    i : INT;
    n : UINT;
END_VAR

(*---IMPL---*)
h := usiActiveClient;
abTx[0] := GVL_IolConst.usiEXT_FUNC_NUM;
abTx[1] := aReq[h].usiPort;
F_IolSetU16BE(ADR(abTx), 2, GVL_IolConst.uiFI_INDEX);
abTx[4] := TO_BYTE(aReq[h].eService);
F_IolSetU16BE(ADR(abTx), 5, aReq[h].uiIndex);
abTx[7] := aReq[h].usiSubindex;
uiTxLen := GVL_IolConst.uiHDR_LEN;
IF aReq[h].eService = E_IolService.WRITE THEN
    n := MIN(aReq[h].uiLen, GVL_IolConst.uiMAX_DATA);
    FOR i := 0 TO UINT_TO_INT(n) - 1 DO
        abTx[GVL_IolConst.uiHDR_LEN + INT_TO_UINT(i)] := aReq[h].abData[i];
    END_FOR
    uiTxLen := GVL_IolConst.uiHDR_LEN + n;
END_IF

// Kiểm khung phản hồi abRx và điền stCur. Layout lỗi (Control 0x80, byte 5..8) là GIẢ ĐỊNH theo spec PNO,
// phải đối chiếu manual AL1100 khi test thật - chỉ cần sửa trong method này.
METHOD PRIVATE ParseResponse : BOOL
VAR
    h : USINT;
    i : INT;
    n : UINT;
END_VAR

(*---IMPL---*)
ParseResponse := FALSE;
h := usiActiveClient;

IF uiRxLen < 5
   OR abRx[0] <> GVL_IolConst.usiEXT_FUNC_NUM
   OR abRx[1] <> aReq[h].usiPort
   OR F_IolGetU16BE(ADR(abRx), 2) <> GVL_IolConst.uiFI_INDEX THEN
    stCur.eErrSource := E_IolErrSource.FRAME;
    RETURN;
END_IF

IF abRx[4] = GVL_IolConst.usiCTRL_ERROR THEN
    IF uiRxLen >= 7 THEN
        stCur.uiIolMasterErr := F_IolGetU16BE(ADR(abRx), 5);
    END_IF
    IF uiRxLen >= 9 THEN
        stCur.uiIolDevErr := F_IolGetU16BE(ADR(abRx), 7);
    END_IF
    IF stCur.uiIolDevErr <> 0 THEN
        stCur.eErrSource := E_IolErrSource.IOL_DEVICE;
    ELSE
        stCur.eErrSource := E_IolErrSource.IOL_MASTER;
    END_IF
    RETURN;
END_IF

IF uiRxLen < GVL_IolConst.uiHDR_LEN
   OR abRx[4] <> TO_BYTE(aReq[h].eService)
   OR F_IolGetU16BE(ADR(abRx), 5) <> aReq[h].uiIndex
   OR abRx[7] <> aReq[h].usiSubindex THEN
    stCur.eErrSource := E_IolErrSource.FRAME;
    RETURN;
END_IF

n := MIN(uiRxLen - GVL_IolConst.uiHDR_LEN, GVL_IolConst.uiMAX_DATA);
FOR i := 0 TO UINT_TO_INT(n) - 1 DO
    stCur.abData[i] := abRx[GVL_IolConst.uiHDR_LEN + INT_TO_UINT(i)];
END_FOR
stCur.uiLen := n;
ParseResponse := TRUE;

// Giao kết quả stCur cho client đang chạy (bỏ nếu client đã Cancel), giải phóng khoá
METHOD PRIVATE Finish
VAR_INPUT
    xErr : BOOL;
END_VAR
VAR
    h : USINT;
END_VAR

(*---IMPL---*)
h := usiActiveClient;
IF h >= 1 AND h <= GVL_IolConst.iQUEUE_SIZE THEN
    stCur.xError := xErr;
    IF NOT axCancel[h] THEN
        aRes[h] := stCur;
        axResReady[h] := TRUE;
    END_IF
    axCancel[h]  := FALSE;
    axPending[h] := FALSE;
END_IF
IF xErr THEN
    udiErrCount := udiErrCount + 1;
ELSE
    udiCallCount := udiCallCount + 1;
END_IF
usiActiveClient := 0;
xWrReq := FALSE;
xRdReq := FALSE;

(*---IMPL---*)
IF usiHandles < INT_TO_USINT(GVL_IolConst.iQUEUE_SIZE) THEN
    usiHandles := usiHandles + 1;
    Register := usiHandles;
ELSE
    Register := 0;
END_IF

// Client gọi 1 lần để nhận handle 1..iQUEUE_SIZE; 0 = hết chỗ
METHOD Register : USINT

// Đưa request của client vào cuối FIFO; FALSE nếu handle sai, đang có request chờ hoặc hàng đợi đầy
METHOD Submit : BOOL
VAR_INPUT
    hHandle : USINT;
END_VAR
VAR_IN_OUT
    stReq : ST_IolRequest;
END_VAR

(*---IMPL---*)
Submit := FALSE;
IF hHandle < 1 OR hHandle > GVL_IolConst.iQUEUE_SIZE THEN
    RETURN;
END_IF
IF axPending[hHandle] OR iCount >= GVL_IolConst.iQUEUE_SIZE THEN
    RETURN;
END_IF
aReq[hHandle] := stReq;
axResReady[hHandle] := FALSE;
axCancel[hHandle]   := FALSE;
axPending[hHandle]  := TRUE;
aQueue[(iHead + iCount) MOD GVL_IolConst.iQUEUE_SIZE] := hHandle;
iCount := iCount + 1;
Submit := TRUE;

// TRUE khi có kết quả cho handle (chép vào stRes và xoá cờ)
METHOD Poll : BOOL
VAR_INPUT
    hHandle : USINT;
END_VAR
VAR_IN_OUT
    stRes : ST_IolResult;
END_VAR

(*---IMPL---*)
Poll := FALSE;
IF hHandle >= 1 AND hHandle <= GVL_IolConst.iQUEUE_SIZE THEN
    IF axResReady[hHandle] THEN
        stRes := aRes[hHandle];
        axResReady[hHandle] := FALSE;
        Poll := TRUE;
    END_IF
END_IF

// Client bỏ request (vd timeout phía client): request còn trong FIFO bị bỏ qua, đang chạy thì huỷ kết quả
METHOD Cancel
VAR_INPUT
    hHandle : USINT;
END_VAR

(*---IMPL---*)
IF hHandle >= 1 AND hHandle <= GVL_IolConst.iQUEUE_SIZE THEN
    IF axPending[hHandle] THEN
        axCancel[hHandle] := TRUE;
    END_IF
    axResReady[hHandle] := FALSE;
END_IF

(* ---- FB_MockRecordAccess.st ---- *)
// Giả lập AL1100 + O5D150 cho CODESYS Simulation: nhận khung IOL_CALL qua Write, trả phản hồi qua Read
// theo layout record CAP 0xB400 (plan mục 4.2). Dữ liệu O5D150 lấy theo IODD; có cờ chèn lỗi để test.
FUNCTION_BLOCK FB_MockRecordAccess IMPLEMENTS ITF_IolRecordAccess
VAR_INPUT
    tDelayWr           : TIME  := T#30MS;     // thời gian giả lập WRREC
    tDelayRd           : TIME  := T#30MS;     // thời gian giả lập RDREC
    usiDevPort         : USINT := GVL_IolConst.usiPORT_O5D150;   // port có O5D150 giả lập
    xDevPresent        : BOOL  := TRUE;       // FALSE -> master trả lỗi truyền thông 0x8004
    usiSimAlign        : USINT := 75;         // giá trị Align (index 69) trả về [%]
    // --- Chèn lỗi ---
    xInjPnioErr        : BOOL;                // WRREC trả STATUS DE80B000
    usiInjBusyCount    : USINT;               // số lần RDREC trả "bận" (B5) cho mỗi request
    uiInjDevErr        : UINT;                // <> 0: mọi request trả lỗi device này (vd 16#8023)
    xInjNoResponse     : BOOL;                // không bao giờ xong -> test timeout
    xInjBadFrame       : BOOL;                // phản hồi byte 0 sai -> lỗi FRAME
    xIdx37NotSupported : BOOL;                // index 37 trả 0x8011 như IODD (không khai báo)
    awInjEvent         : ARRAY[0..3] OF WORD; // thêm event bất kỳ vào danh sách index 37 (0 = trống)
END_VAR
VAR_OUTPUT
    udiWrCount    : UDINT;
    udiRdCount    : UDINT;
    usiLastSysCmd : USINT;                    // System Command gần nhất nhận được
    xEvt1Active   : BOOL;                     // Test Event 0x8DFE đang active
    xEvt2Active   : BOOL;                     // Test Event 0x8DFF đang active
END_VAR
VAR
    xInit       : BOOL;
    aStore      : ARRAY[0..19] OF ST_MockParam;
    iStoreCount : INT;
    tonWr       : TON;
    tonRd       : TON;
    xWrActive   : BOOL;
    xWrFinished : BOOL;
    xWrFailed   : BOOL;
    dwWrStat    : DWORD;
    xRdActive   : BOOL;
    xRdFinished : BOOL;
    xRdFailed   : BOOL;
    dwRdStat    : DWORD;
    iRdLenOut   : INT;
    abReq       : ARRAY[0..GVL_IolConst.uiMAX_REC - 1] OF BYTE;
    uiReqLen    : UINT;
    abResp      : ARRAY[0..GVL_IolConst.uiMAX_REC - 1] OF BYTE;
    uiRespLen   : UINT;
    xRespReady  : BOOL;
    usiBusyLeft : USINT;
    abTmp       : ARRAY[0..63] OF BYTE;
END_VAR

(*---IMPL---*)
// Không có xử lý chu kỳ: Write/Read do FB_IolMaster gọi mỗi chu kỳ.
IF NOT xInit THEN
    InitStore();
END_IF

METHOD Write : BOOL
VAR_INPUT
    xReq   : BOOL;
    dwId   : DWORD;
    iIndex : INT;
    iLen   : INT;
    pData  : POINTER TO BYTE;
END_VAR
VAR_OUTPUT
    xDone    : BOOL;
    xBusy    : BOOL;
    xError   : BOOL;
    dwStatus : DWORD;
END_VAR
VAR
    i : INT;
END_VAR

(*---IMPL---*)
IF NOT xInit THEN
    InitStore();
END_IF

IF NOT xReq THEN
    // REQ hạ: sẵn sàng cho request mới
    xWrActive   := FALSE;
    xWrFinished := FALSE;
    xWrFailed   := FALSE;
    tonWr(IN := FALSE);
ELSIF NOT xWrActive AND NOT xWrFinished THEN
    // sườn lên REQ: chụp khung request
    uiReqLen := INT_TO_UINT(LIMIT(0, iLen, UINT_TO_INT(GVL_IolConst.uiMAX_REC)));
    IF pData = 0 THEN
        uiReqLen := 0;
    END_IF
    FOR i := 0 TO UINT_TO_INT(uiReqLen) - 1 DO
        abReq[i] := pData[i];
    END_FOR
    xWrActive := TRUE;
END_IF

IF xWrActive THEN
    tonWr(IN := TRUE, PT := tDelayWr);
    IF tonWr.Q AND NOT xInjNoResponse THEN
        tonWr(IN := FALSE);
        xWrActive   := FALSE;
        xWrFinished := TRUE;
        udiWrCount  := udiWrCount + 1;
        IF xInjPnioErr OR iIndex <> UINT_TO_INT(GVL_IolConst.uiCAP_INDEX) THEN
            xWrFailed := TRUE;
            dwWrStat  := 16#DE80B000;          // invalid index
        ELSE
            xWrFailed := FALSE;
            dwWrStat  := 0;
            ProcessRequest();
        END_IF
    END_IF
END_IF

xBusy  := xWrActive;
xDone  := xWrFinished AND NOT xWrFailed;
xError := xWrFinished AND xWrFailed;
IF xError THEN
    dwStatus := dwWrStat;
ELSE
    dwStatus := 0;
END_IF
Write := xWrFinished;

METHOD Read : BOOL
VAR_INPUT
    xReq   : BOOL;
    dwId   : DWORD;
    iIndex : INT;
    iMLen  : INT;
    pData  : POINTER TO BYTE;
END_VAR
VAR_OUTPUT
    xValid   : BOOL;
    xBusy    : BOOL;
    xError   : BOOL;
    dwStatus : DWORD;
    iLen     : INT;
END_VAR
VAR
    i : INT;
    n : INT;
END_VAR

(*---IMPL---*)
IF NOT xInit THEN
    InitStore();
END_IF

IF NOT xReq THEN
    xRdActive   := FALSE;
    xRdFinished := FALSE;
    xRdFailed   := FALSE;
    tonRd(IN := FALSE);
ELSIF NOT xRdActive AND NOT xRdFinished THEN
    xRdActive := TRUE;
END_IF

IF xRdActive THEN
    tonRd(IN := TRUE, PT := tDelayRd);
    IF tonRd.Q AND NOT xInjNoResponse THEN
        tonRd(IN := FALSE);
        xRdActive   := FALSE;
        xRdFinished := TRUE;
        udiRdCount  := udiRdCount + 1;
        iRdLenOut   := 0;
        IF iIndex <> UINT_TO_INT(GVL_IolConst.uiCAP_INDEX) THEN
            xRdFailed := TRUE;
            dwRdStat  := 16#DE80B000;          // invalid index
        ELSIF usiBusyLeft > 0 OR NOT xRespReady THEN
            // master chưa xử lý xong ISDU (hoặc chưa có request) -> state conflict, client retry
            IF usiBusyLeft > 0 THEN
                usiBusyLeft := usiBusyLeft - 1;
            END_IF
            xRdFailed := TRUE;
            dwRdStat  := 16#DE80B500;
        ELSE
            n := MIN(UINT_TO_INT(uiRespLen), iMLen);
            IF pData = 0 THEN
                n := 0;
            END_IF
            FOR i := 0 TO n - 1 DO
                pData[i] := abResp[i];
            END_FOR
            iRdLenOut  := n;
            xRespReady := FALSE;               // phản hồi chỉ đọc được 1 lần
            xRdFailed  := FALSE;
            dwRdStat   := 0;
        END_IF
    END_IF
END_IF

xBusy  := xRdActive;
xValid := xRdFinished AND NOT xRdFailed;
xError := xRdFinished AND xRdFailed;
IF xError THEN
    dwStatus := dwRdStat;
ELSE
    dwStatus := 0;
END_IF
IF xValid THEN
    iLen := iRdLenOut;
ELSE
    iLen := 0;
END_IF
Read := xRdFinished;

(*---IMPL---*)
iStoreCount := 0;
// --- Nhận dạng chuẩn 16..24 ---
AddStr(16,  E_IolAccess.RO, 'ifm electronic gmbh');
AddStr(17,  E_IolAccess.RO, 'www.ifm.com');
AddStr(18,  E_IolAccess.RO, 'O5D150');
AddStr(19,  E_IolAccess.RO, 'O5D150');
AddStr(20,  E_IolAccess.RO, 'Laser distance sensor (SIM)');
AddStr(21,  E_IolAccess.RO, 'SIM0001');
AddStr(22,  E_IolAccess.RO, 'AB');
AddStr(23,  E_IolAccess.RO, 'SIM 1.0');
AddStr(24,  E_IolAccess.RW, '***');
// --- Tham số theo IODD (giá trị big-endian) ---
AddRaw(60,  E_IolAccess.RW, 4, 16#00640000);   // SP1 = 100 cm, SP2 = 0 (not used)
AddRaw(61,  E_IolAccess.RW, 4, 16#00010000);   // Logic = 0 NO, Mode = 1, Hyst = 0
AddRaw(64,  E_IolAccess.RO, 4, 16#000500C8);   // Limit min 5 cm, max 200 cm
AddRaw(69,  E_IolAccess.RO, 1, 75);            // Align %
AddRaw(74,  E_IolAccess.RW, 2, 0);             // dFO
AddRaw(76,  E_IolAccess.RW, 2, 0);             // dS
AddRaw(78,  E_IolAccess.RW, 2, 0);             // dr
AddRaw(80,  E_IolAccess.RW, 1, 1);             // Laser On
AddRaw(96,  E_IolAccess.RW, 1, 1);             // Display On
AddRaw(100, E_IolAccess.RW, 1, 1);             // KeyLock Unlocked
xInit := TRUE;

// Nạp bảng dữ liệu O5D150 mặc định (cũng dùng cho System Command 130 factory reset)
METHOD PRIVATE InitStore

// Thêm 1 index số (1, 2 hoặc 4 byte, big-endian) vào bảng giả lập
METHOD PRIVATE AddRaw
VAR_INPUT
    uiIndex : UINT;
    eAccess : E_IolAccess;
    uiLen   : UINT;          // 1, 2 hoặc 4
    dwVal   : DWORD;
END_VAR

(*---IMPL---*)
IF iStoreCount > 19 THEN
    RETURN;
END_IF
aStore[iStoreCount].uiIndex := uiIndex;
aStore[iStoreCount].eAccess := eAccess;
aStore[iStoreCount].uiLen   := uiLen;
CASE uiLen OF
    1: aStore[iStoreCount].abData[0] := DWORD_TO_BYTE(dwVal);
    2: F_IolSetU16BE(ADR(aStore[iStoreCount].abData), 0, DWORD_TO_UINT(dwVal));
ELSE
    aStore[iStoreCount].uiLen := 4;
    F_IolSetU32BE(ADR(aStore[iStoreCount].abData), 0, dwVal);
END_CASE
iStoreCount := iStoreCount + 1;

// Thêm 1 index chuỗi (StringT, không ký tự kết thúc) vào bảng giả lập
METHOD PRIVATE AddStr
VAR_INPUT
    uiIndex : UINT;
    eAccess : E_IolAccess;
    sVal    : STRING(63);
END_VAR
VAR
    pSrc : POINTER TO BYTE;
    n    : INT;
    i    : INT;
END_VAR

(*---IMPL---*)
IF iStoreCount > 19 THEN
    RETURN;
END_IF
pSrc := ADR(sVal);
n := LEN(sVal);
aStore[iStoreCount].uiIndex := uiIndex;
aStore[iStoreCount].eAccess := eAccess;
aStore[iStoreCount].uiLen   := INT_TO_UINT(n);
FOR i := 0 TO n - 1 DO
    aStore[iStoreCount].abData[i] := pSrc[i];
END_FOR
iStoreCount := iStoreCount + 1;

// Vị trí index trong bảng, -1 nếu không có
METHOD PRIVATE FindStore : INT
VAR_INPUT
    uiIndex : UINT;
END_VAR
VAR
    i : INT;
END_VAR

(*---IMPL---*)
FindStore := -1;
FOR i := 0 TO iStoreCount - 1 DO
    IF aStore[i].uiIndex = uiIndex THEN
        FindStore := i;
        RETURN;
    END_IF
END_FOR

// Vị trí byte của subindex trong record (theo IODD O5D150); FALSE = subindex không tồn tại
METHOD PRIVATE SubRange : BOOL
VAR_INPUT
    iStore  : INT;
    usiSub  : USINT;
END_VAR
VAR_OUTPUT
    uiOff : UINT;
    uiLen : UINT;
END_VAR

(*---IMPL---*)
SubRange := TRUE;
uiOff := 0;
uiLen := 0;
IF usiSub = 0 THEN
    uiLen := aStore[iStore].uiLen;
    RETURN;
END_IF
CASE aStore[iStore].uiIndex OF
    60:                                   // SP: sub1 SP1, sub2 SP2
        CASE usiSub OF
            1: uiOff := 0; uiLen := 2;
            2: uiOff := 2; uiLen := 2;
        ELSE
            SubRange := FALSE;
        END_CASE
    61:                                   // Config: sub1 Logic, sub2 Mode, sub3 Hyst
        CASE usiSub OF
            1: uiOff := 0; uiLen := 1;
            2: uiOff := 1; uiLen := 1;
            3: uiOff := 2; uiLen := 2;
        ELSE
            SubRange := FALSE;
        END_CASE
    64:                                   // Limit: sub1 min, sub2 max
        CASE usiSub OF
            1: uiOff := 0; uiLen := 2;
            2: uiOff := 2; uiLen := 2;
        ELSE
            SubRange := FALSE;
        END_CASE
ELSE
    SubRange := FALSE;
END_CASE

// Kiểm dải giá trị của cả record sau khi ghi (theo IODD); FALSE -> device trả 0x8030
METHOD PRIVATE CheckImage : BOOL
VAR_INPUT
    uiIndex : UINT;
    pImg    : POINTER TO BYTE;
END_VAR
VAR
    uiV1 : UINT;
    uiV2 : UINT;
END_VAR

(*---IMPL---*)
CheckImage := TRUE;
CASE uiIndex OF
    60:                                         // SP1 5..200 cm, SP2 = 0 (not used)
        uiV1 := F_IolGetU16BE(pImg, 0);
        uiV2 := F_IolGetU16BE(pImg, 2);
        CheckImage := (uiV1 >= 5) AND (uiV1 <= 200) AND (uiV2 = 0);
    61:                                         // Logic 0..1, Mode = 1, Hyst = 0
        CheckImage := (pImg[0] <= 1) AND (pImg[1] = 1) AND (F_IolGetU16BE(pImg, 2) = 0);
    74, 76, 78:                                 // dFO / dS / dr 0..2000
        CheckImage := F_IolGetU16BE(pImg, 0) <= 2000;
    80, 100:                                    // Laser, KeyLock 0..1
        CheckImage := pImg[0] <= 1;
    96:                                         // Display 0..2
        CheckImage := pImg[0] <= 2;
END_CASE

// Hoàn tất phản hồi OK: header đã echo trong abResp[0..7], dữ liệu đọc ở abResp[8..]
METHOD PRIVATE RespOk
VAR_INPUT
    uiDataLen : UINT;
END_VAR

(*---IMPL---*)
uiRespLen := GVL_IolConst.uiHDR_LEN + uiDataLen;
IF xInjBadFrame THEN
    abResp[0] := 0;
END_IF

// Phản hồi lỗi: Control = 0x80, byte 5..6 IOL_M_ErrorCode, byte 7..8 IOL_D_ErrorCode (layout giả định plan 4.2)
METHOD PRIVATE RespErr
VAR_INPUT
    uiMasterErr : UINT;
    uiDevErr    : UINT;
END_VAR

(*---IMPL---*)
abResp[4] := GVL_IolConst.usiCTRL_ERROR;
F_IolSetU16BE(ADR(abResp), 5, uiMasterErr);
F_IolSetU16BE(ADR(abResp), 7, uiDevErr);
uiRespLen := 9;
IF xInjBadFrame THEN
    abResp[0] := 0;
END_IF

// Xử lý 1 khung IOL_CALL đã nhận (abReq), tạo phản hồi trong abResp như AL1100 + O5D150
METHOD PRIVATE ProcessRequest
VAR
    usiPort   : USINT;
    bCtrl     : BYTE;
    uiIdx     : UINT;
    usiSub    : USINT;
    uiDataLen : UINT;
    iS        : INT;
    uiOff     : UINT;
    uiSubLen  : UINT;
    i         : INT;
    n         : UINT;
    awList    : ARRAY[0..5] OF WORD;   // event đang active để trả ở index 37
    abQual    : ARRAY[0..5] OF BYTE;
END_VAR

(*---IMPL---*)
xRespReady  := TRUE;
usiBusyLeft := usiInjBusyCount;
FOR i := 0 TO 7 DO                       // phản hồi echo header request
    abResp[i] := abReq[i];
END_FOR

// ---------- 1. Kiểm khung ----------
IF uiReqLen < GVL_IolConst.uiHDR_LEN
   OR abReq[0] <> GVL_IolConst.usiEXT_FUNC_NUM
   OR F_IolGetU16BE(ADR(abReq), 2) <> GVL_IolConst.uiFI_INDEX THEN
    RespErr(16#7001, 0);                 // wrong IOL_CALL
    RETURN;
END_IF
usiPort   := abReq[1];
bCtrl     := abReq[4];
uiIdx     := F_IolGetU16BE(ADR(abReq), 5);
usiSub    := abReq[7];
uiDataLen := uiReqLen - GVL_IolConst.uiHDR_LEN;

IF usiPort < 1 OR usiPort > 4 THEN
    RespErr(16#8001, 0);                 // port không hợp lệ
    RETURN;
END_IF
IF usiPort <> usiDevPort OR NOT xDevPresent THEN
    RespErr(16#8004, 0);                 // không liên lạc được device trên port
    RETURN;
END_IF
IF bCtrl <> GVL_IolConst.usiCTRL_READ AND bCtrl <> GVL_IolConst.usiCTRL_WRITE THEN
    RespErr(16#7001, 0);
    RETURN;
END_IF
IF uiInjDevErr <> 0 THEN
    RespErr(0, uiInjDevErr);
    RETURN;
END_IF

// ---------- 2. Index 37: Detailed Device Status (3 byte/entry: qualifier + code) ----------
IF uiIdx = GVL_O5D150_Def.uiIDX_EVT_LIST THEN
    IF bCtrl = GVL_IolConst.usiCTRL_WRITE THEN
        RespErr(0, GVL_IolConst.uiERR_ACCESS);
    ELSIF xIdx37NotSupported THEN
        RespErr(0, GVL_IolConst.uiERR_IDX_NA);
    ELSE
        awList[0] := SEL(xEvt1Active, 0, 16#8DFE);  abQual[0] := 16#D4;   // appear, notification, device, application
        awList[1] := SEL(xEvt2Active, 0, 16#8DFF);  abQual[1] := 16#D4;
        FOR i := 0 TO 3 DO
            awList[i + 2] := awInjEvent[i];
            abQual[i + 2] := 16#E4;                                        // appear, warning
        END_FOR
        n := 0;
        FOR i := 0 TO 5 DO
            IF awList[i] <> 0 THEN
                abResp[8 + n] := abQual[i];
                F_IolSetU16BE(ADR(abResp), 9 + n, WORD_TO_UINT(awList[i]));
                n := n + 3;
            END_IF
        END_FOR
        RespOk(n);
    END_IF
    RETURN;
END_IF

// ---------- 3. Index 2: System Command ----------
IF uiIdx = GVL_O5D150_Def.uiIDX_SYS_CMD THEN
    IF bCtrl = GVL_IolConst.usiCTRL_READ THEN
        RespErr(0, GVL_IolConst.uiERR_ACCESS);      // write only
    ELSIF uiDataLen > 1 THEN
        RespErr(0, 16#8033);
    ELSIF uiDataLen < 1 THEN
        RespErr(0, 16#8034);
    ELSE
        usiLastSysCmd := abReq[8];
        CASE usiLastSysCmd OF
            130: InitStore(); xEvt1Active := FALSE; xEvt2Active := FALSE; RespOk(0);
            240: xEvt1Active := TRUE;  RespOk(0);
            241: xEvt1Active := FALSE; RespOk(0);
            242: xEvt2Active := TRUE;  RespOk(0);
            243: xEvt2Active := FALSE; RespOk(0);
        ELSE
            RespErr(0, 16#8035);                    // lệnh không có trong IODD
        END_CASE
    END_IF
    RETURN;
END_IF

// ---------- 4. Bảng tham số ----------
iS := FindStore(uiIdx);
IF iS < 0 THEN
    RespErr(0, GVL_IolConst.uiERR_IDX_NA);
    RETURN;
END_IF
IF NOT SubRange(iStore := iS, usiSub := usiSub, uiOff => uiOff, uiLen => uiSubLen) THEN
    RespErr(0, GVL_IolConst.uiERR_SUBIDX_NA);
    RETURN;
END_IF

IF bCtrl = GVL_IolConst.usiCTRL_READ THEN
    IF aStore[iS].eAccess = E_IolAccess.WO THEN
        RespErr(0, GVL_IolConst.uiERR_ACCESS);
        RETURN;
    END_IF
    IF uiIdx = 69 THEN
        aStore[iS].abData[0] := usiSimAlign;
    END_IF
    FOR i := 0 TO UINT_TO_INT(uiSubLen) - 1 DO
        abResp[8 + i] := aStore[iS].abData[uiOff + INT_TO_UINT(i)];
    END_FOR
    RespOk(uiSubLen);
ELSE
    IF aStore[iS].eAccess = E_IolAccess.RO THEN
        RespErr(0, GVL_IolConst.uiERR_ACCESS);
    ELSIF uiDataLen > uiSubLen THEN
        RespErr(0, 16#8033);
    ELSIF uiDataLen < uiSubLen THEN
        RespErr(0, 16#8034);
    ELSE
        // ghép giá trị mới vào bản sao record rồi kiểm dải trước khi chấp nhận
        abTmp := aStore[iS].abData;
        FOR i := 0 TO UINT_TO_INT(uiSubLen) - 1 DO
            abTmp[uiOff + INT_TO_UINT(i)] := abReq[8 + i];
        END_FOR
        IF CheckImage(uiIdx, ADR(abTmp)) THEN
            aStore[iS].abData := abTmp;
            RespOk(0);
        ELSE
            RespErr(0, GVL_IolConst.uiERR_RANGE);
        END_IF
    END_IF
END_IF

(* ---- FB_PnRecordAccess.st ---- *)
// Transport PROFINET thật: bọc CommFB.WRREC / CommFB.RDREC tới submodule CAP của AL1100.
// HIỆN LÀ KHUNG: chưa có PN Controller + AL1100 được duyệt (IP, station name, license) nên chưa gọi CommFB;
// mọi request trả lỗi dwSTAT_NOT_CONFIGURED để master báo rõ thay vì treo.
// TODO PROFINET:
//   1. Thêm AL1100 dưới PN_Controller, đặt bus cycle task = MainTask.
//   2. VAR: fbWr : CommFB.WRREC; fbRd : CommFB.RDREC;
//   3. dwId := CommFB.SUBSLOT_ID(EN := TRUE, ID := <AL1100>.DeviceID, SLOT := usiSlot, SUBSLOT := usiSubslot);
//      dwId = CommFB.Constants.INVALID_ID -> lỗi cấu hình.
//   4. Write: fbWr(REQ := xReq, ID := dwId, INDEX := iIndex, LEN := iLen, RECORD := <buffer>); xDone := fbWr.DONE ...
//      Read : fbRd(REQ := xReq, ID := dwId, INDEX := iIndex, MLEN := iMLen, RECORD := <buffer>); xValid := fbRd.VALID; iLen := fbRd.LEN ...
//      Kiểu chân RECORD (ANY / POINTER) phải xem trong Library Manager rồi copy buffer cho đúng.
//   5. Luôn viết đủ namespace CommFB.* (tránh trùng tên với lib Turck commfb*).
FUNCTION_BLOCK FB_PnRecordAccess IMPLEMENTS ITF_IolRecordAccess
VAR_INPUT
    usiSlot    : USINT := GVL_IolConst.usiAL1_SLOT;
    usiSubslot : USINT := GVL_IolConst.usiAL1_SUBSLOT_CAP;
END_VAR
VAR_OUTPUT
    xNotConfigured : BOOL := TRUE;    // TRUE khi FB còn là khung
END_VAR

(*---IMPL---*)
// Không có xử lý chu kỳ: toàn bộ việc nằm trong method Write/Read (gọi bởi FB_IolMaster).
xNotConfigured := TRUE;

METHOD Write : BOOL
VAR_INPUT
    xReq   : BOOL;
    dwId   : DWORD;
    iIndex : INT;
    iLen   : INT;
    pData  : POINTER TO BYTE;
END_VAR
VAR_OUTPUT
    xDone    : BOOL;
    xBusy    : BOOL;
    xError   : BOOL;
    dwStatus : DWORD;
END_VAR

(*---IMPL---*)
// TODO PROFINET: thay bằng CommFB.WRREC (xem ghi chú khai báo FB)
xDone  := FALSE;
xBusy  := FALSE;
xError := xReq;
IF xReq THEN
    dwStatus := GVL_IolConst.dwSTAT_NOT_CONFIGURED;
ELSE
    dwStatus := 0;
END_IF
Write := xReq;

METHOD Read : BOOL
VAR_INPUT
    xReq   : BOOL;
    dwId   : DWORD;
    iIndex : INT;
    iMLen  : INT;
    pData  : POINTER TO BYTE;
END_VAR
VAR_OUTPUT
    xValid   : BOOL;
    xBusy    : BOOL;
    xError   : BOOL;
    dwStatus : DWORD;
    iLen     : INT;
END_VAR

(*---IMPL---*)
// TODO PROFINET: thay bằng CommFB.RDREC (xem ghi chú khai báo FB)
xValid := FALSE;
xBusy  := FALSE;
xError := xReq;
iLen   := 0;
IF xReq THEN
    dwStatus := GVL_IolConst.dwSTAT_NOT_CONFIGURED;
ELSE
    dwStatus := 0;
END_IF
Read := xReq;

(* ---- PLC_PRG.st ---- *)
PROGRAM PLC_PRG
VAR
    fbSeq    : FB_OutSeq;     // bộ tạo trình tự ngõ ra
    xRunReq  : BOOL;          // chốt Start/Stop
    byManual : BYTE;          // ảnh ngõ ra tay
    i        : INT;
END_VAR

(*---IMPL---*)
// ---------- 1. Start / Stop (Stop ưu tiên) ----------
IF GVL_HMI.xCmdStop THEN
    xRunReq := FALSE;
ELSIF GVL_HMI.xCmdStart THEN
    xRunReq := TRUE;
END_IF
GVL_HMI.xCmdStart := FALSE;
GVL_HMI.xCmdStop  := FALSE;

// ---------- 2. Giới hạn thông số từ visu ----------
GVL_HMI.iModeSel  := LIMIT(0, GVL_HMI.iModeSel, 13);
GVL_HMI.udiStepMs := LIMIT(50, GVL_HMI.udiStepMs, 2000);
GVL_HMI.udiDemoS  := LIMIT(2, GVL_HMI.udiDemoS, 60);

byManual := 0;
FOR i := 0 TO 7 DO
    IF GVL_HMI.axManual[i] THEN
        byManual := byManual OR SHL(BYTE#1, i);
    END_IF
END_FOR

// ---------- 3. Tạo trình tự (MANUAL chạy không cần Start) ----------
fbSeq(
    xRun      := (xRunReq AND GVL_HMI.iModeSel <> E_SeqMode.OFF) OR GVL_HMI.iModeSel = E_SeqMode.MANUAL,
    eMode     := GVL_HMI.iModeSel,
    tStep     := UDINT_TO_TIME(GVL_HMI.udiStepMs),
    tDemoHold := UDINT_TO_TIME(GVL_HMI.udiDemoS * 1000),
    xReverse  := GVL_HMI.xReverse,
    byManual  := byManual);

// ---------- 4. Ghi ngõ ra DXP ----------
GVL_IO.xQ_Ch8  := fbSeq.byOut.0;
GVL_IO.xQ_Ch9  := fbSeq.byOut.1;
GVL_IO.xQ_Ch10 := fbSeq.byOut.2;
GVL_IO.xQ_Ch11 := fbSeq.byOut.3;
GVL_IO.xQ_Ch12 := fbSeq.byOut.4;
GVL_IO.xQ_Ch13 := fbSeq.byOut.5;
GVL_IO.xQ_Ch14 := fbSeq.byOut.6;
GVL_IO.xQ_Ch15 := fbSeq.byOut.7;

// ---------- 5. Trạng thái lên visu ----------
GVL_HMI.xRunning    := fbSeq.xRun;
GVL_HMI.byOut       := fbSeq.byOut;
GVL_HMI.uiStep      := fbSeq.uiStep;
GVL_HMI.iModeActive := fbSeq.eActive;
FOR i := 0 TO 7 DO
    GVL_HMI.axOut[i] := (SHR(fbSeq.byOut, i) AND 1) <> 0;
END_FOR
FOR i := 0 TO 13 DO
    GVL_HMI.axModeSel[i] := (GVL_HMI.iModeSel = i);
END_FOR
GVL_HMI.xNotManual := (GVL_HMI.iModeSel <> E_SeqMode.MANUAL);
GVL_HMI.axFb[0] := GVL_IO.xI_Ch8;
GVL_HMI.axFb[1] := GVL_IO.xI_Ch9;
GVL_HMI.axFb[2] := GVL_IO.xI_Ch10;
GVL_HMI.axFb[3] := GVL_IO.xI_Ch11;
GVL_HMI.axFb[4] := GVL_IO.xI_Ch12;
GVL_HMI.axFb[5] := GVL_IO.xI_Ch13;
GVL_HMI.axFb[6] := GVL_IO.xI_Ch14;
GVL_HMI.axFb[7] := GVL_IO.xI_Ch15;

CASE fbSeq.eActive OF
    E_SeqMode.OFF:       GVL_HMI.sModeName := "OFF - Tắt";
    E_SeqMode.CHASE:     GVL_HMI.sModeName := "Chạy đuổi";
    E_SeqMode.PINGPONG:  GVL_HMI.sModeName := "Qua lại";
    E_SeqMode.FILL:      GVL_HMI.sModeName := "Sáng dồn / tắt dần";
    E_SeqMode.STACK:     GVL_HMI.sModeName := "Xếp chồng";
    E_SeqMode.BLINK:     GVL_HMI.sModeName := "Nhấp nháy";
    E_SeqMode.ALTERNATE: GVL_HMI.sModeName := "Chẵn / lẻ";
    E_SeqMode.BINARY:    GVL_HMI.sModeName := "Đếm nhị phân";
    E_SeqMode.CENTER:    GVL_HMI.sModeName := "Từ giữa ra";
    E_SeqMode.WAVE:      GVL_HMI.sModeName := "Sóng 3 đèn";
    E_SeqMode.PAIR:      GVL_HMI.sModeName := "Cặp đèn";
    E_SeqMode.RANDOM:    GVL_HMI.sModeName := "Ngẫu nhiên";
    E_SeqMode.MANUAL:    GVL_HMI.sModeName := "Bật tay";
END_CASE

// ---------- 6. IO-Link AL1100 / O5D150 ----------
PRG_IOLink();
